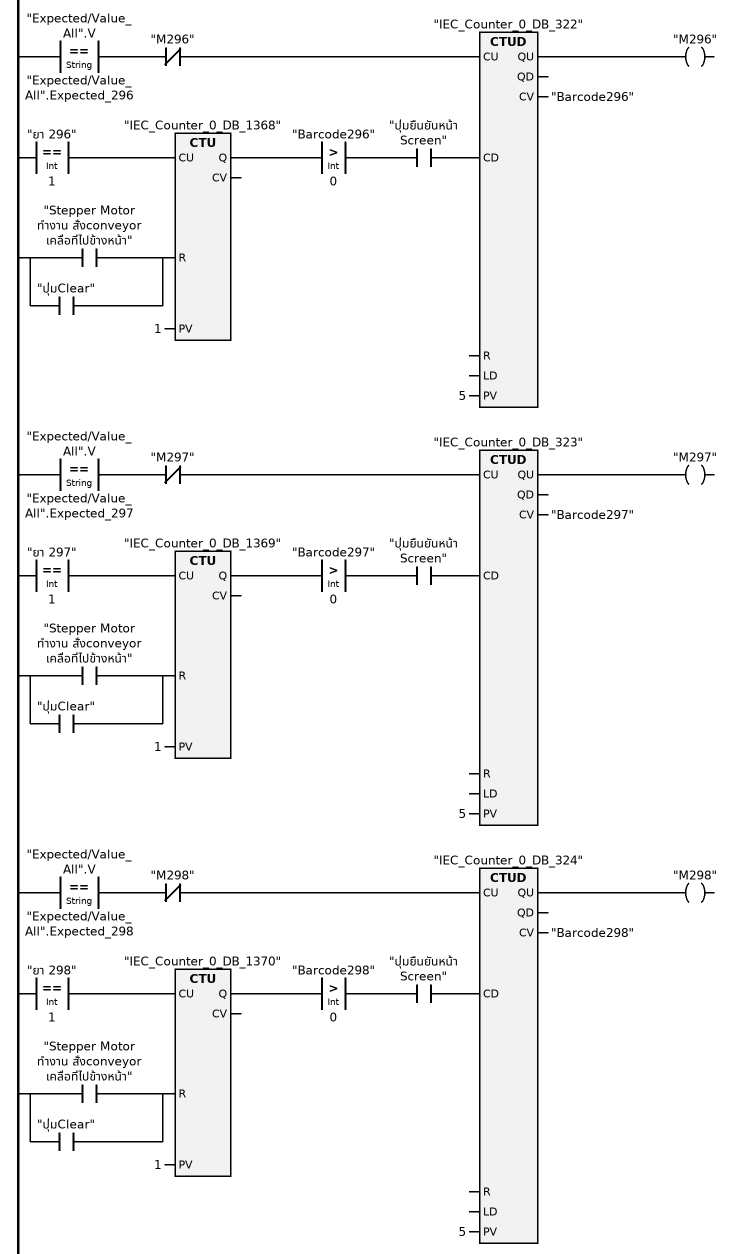
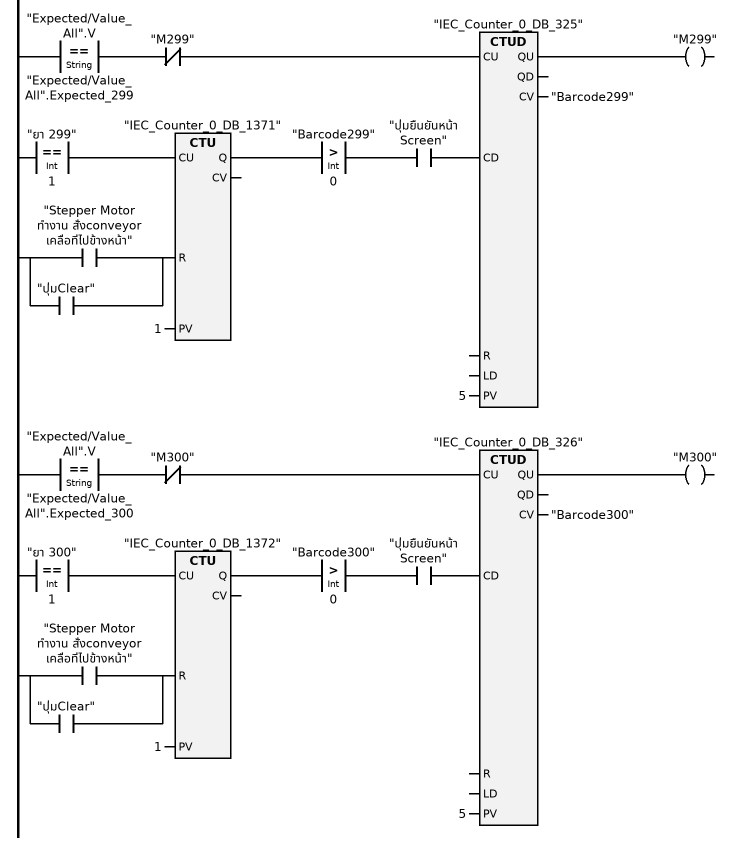
   "IEC_Counter_0_DB_1353".CTU(CU := "ยา 281" = 1,
                           R := "Stepper Motor ทำงาน สั่งconveyor เคลื่อที่ไปข้างหน้า" OR "ปุ่มClear",
                           PV := 1);
   "IEC_Counter_0_DB_307".CTUD(CU := ("Expected/Value_All".V = "Expected/Value_All".Expected_281) AND NOT "M281",
                           CD := "IEC_Counter_0_DB_1353".Q AND ("Barcode281" > 0) AND "ปุ่มยืนยันหน้า Screen",
                           PV := 5,
                           CV => "Barcode281");
   "M281" := "IEC_Counter_0_DB_307".QU;
   "IEC_Counter_0_DB_1354".CTU(CU := "ยา 282" = 1,
                           R := "Stepper Motor ทำงาน สั่งconveyor เคลื่อที่ไปข้างหน้า" OR "ปุ่มClear",
                           PV := 1);
   "IEC_Counter_0_DB_308".CTUD(CU := ("Expected/Value_All".V = "Expected/Value_All".Expected_282) AND NOT "M282",
                           CD := "IEC_Counter_0_DB_1354".Q AND ("Barcode282" > 0) AND "ปุ่มยืนยันหน้า Screen",
                           PV := 5,
                           CV => "Barcode282");
   "M282" := "IEC_Counter_0_DB_308".QU;
   "IEC_Counter_0_DB_1355".CTU(CU := "ยา 283" = 1,
                           R := "Stepper Motor ทำงาน สั่งconveyor เคลื่อที่ไปข้างหน้า" OR "ปุ่มClear",
                           PV := 1);
   "IEC_Counter_0_DB_309".CTUD(CU := ("Expected/Value_All".V = "Expected/Value_All".Expected_283) AND NOT "M283",
                           CD := "IEC_Counter_0_DB_1355".Q AND ("Barcode283" > 0) AND "ปุ่มยืนยันหน้า Screen",
                           PV := 5,
                           CV => "Barcode283");
   "M283" := "IEC_Counter_0_DB_309".QU;
   "IEC_Counter_0_DB_1356".CTU(CU := "ยา 284" = 1,
                           R := "Stepper Motor ทำงาน สั่งconveyor เคลื่อที่ไปข้างหน้า" OR "ปุ่มClear",
                           PV := 1);
   "IEC_Counter_0_DB_310".CTUD(CU := ("Expected/Value_All".V = "Expected/Value_All".Expected_284) AND NOT "M284",
                           CD := "IEC_Counter_0_DB_1356".Q AND ("Barcode284" > 0) AND "ปุ่มยืนยันหน้า Screen",
                           PV := 5,
                           CV => "Barcode284");
   "M284" := "IEC_Counter_0_DB_310".QU;
   "IEC_Counter_0_DB_1357".CTU(CU := "ยา 285" = 1,
                           R := "Stepper Motor ทำงาน สั่งconveyor เคลื่อที่ไปข้างหน้า" OR "ปุ่มClear",
                           PV := 1);
   "IEC_Counter_0_DB_311".CTUD(CU := ("Expected/Value_All".V = "Expected/Value_All".Expected_285) AND NOT "M285",
                           CD := "IEC_Counter_0_DB_1357".Q AND ("Barcode285" > 0) AND "ปุ่มยืนยันหน้า Screen",
                           PV := 5,
                           CV => "Barcode285");
   "M285" := "IEC_Counter_0_DB_311".QU;
   "IEC_Counter_0_DB_1358".CTU(CU := "ยา 286" = 1,
                           R := "Stepper Motor ทำงาน สั่งconveyor เคลื่อที่ไปข้างหน้า" OR "ปุ่มClear",
                           PV := 1);
   "IEC_Counter_0_DB_312".CTUD(CU := ("Expected/Value_All".V = "Expected/Value_All".Expected_286) AND NOT "M286",
                           CD := "IEC_Counter_0_DB_1358".Q AND ("Barcode286" > 0) AND "ปุ่มยืนยันหน้า Screen",
                           PV := 5,
                           CV => "Barcode286");
   "M286" := "IEC_Counter_0_DB_312".QU;
   "IEC_Counter_0_DB_1359".CTU(CU := "ยา 287" = 1,
                           R := "Stepper Motor ทำงาน สั่งconveyor เคลื่อที่ไปข้างหน้า" OR "ปุ่มClear",
                           PV := 1);
   "IEC_Counter_0_DB_313".CTUD(CU := ("Expected/Value_All".V = "Expected/Value_All".Expected_287) AND NOT "M287",
                           CD := "IEC_Counter_0_DB_1359".Q AND ("Barcode287" > 0) AND "ปุ่มยืนยันหน้า Screen",
                           PV := 5,
                           CV => "Barcode287");
   "M287" := "IEC_Counter_0_DB_313".QU;
   "IEC_Counter_0_DB_1360".CTU(CU := "ยา 288" = 1,
                           R := "Stepper Motor ทำงาน สั่งconveyor เคลื่อที่ไปข้างหน้า" OR "ปุ่มClear",
                           PV := 1);
   "IEC_Counter_0_DB_314".CTUD(CU := ("Expected/Value_All".V = "Expected/Value_All".Expected_288) AND NOT "M288",
                           CD := "IEC_Counter_0_DB_1360".Q AND ("Barcode288" > 0) AND "ปุ่มยืนยันหน้า Screen",
                           PV := 5,
                           CV => "Barcode288");
   "M288" := "IEC_Counter_0_DB_314".QU;
   "IEC_Counter_0_DB_1361".CTU(CU := "ยา 289" = 1,
                           R := "Stepper Motor ทำงาน สั่งconveyor เคลื่อที่ไปข้างหน้า" OR "ปุ่มClear",
                           PV := 1);
   "IEC_Counter_0_DB_315".CTUD(CU := ("Expected/Value_All".V = "Expected/Value_All".Expected_289) AND NOT "M289",
                           CD := "IEC_Counter_0_DB_1361".Q AND ("Barcode289" > 0) AND "ปุ่มยืนยันหน้า Screen",
                           PV := 5,
                           CV => "Barcode289");
   "M289" := "IEC_Counter_0_DB_315".QU;
   "IEC_Counter_0_DB_1362".CTU(CU := "ยา 290" = 1,
                           R := "Stepper Motor ทำงาน สั่งconveyor เคลื่อที่ไปข้างหน้า" OR "ปุ่มClear",
                           PV := 1);
   "IEC_Counter_0_DB_316".CTUD(CU := ("Expected/Value_All".V = "Expected/Value_All".Expected_290) AND NOT "M290",
                           CD := "IEC_Counter_0_DB_1362".Q AND ("Barcode290" > 0) AND "ปุ่มยืนยันหน้า Screen",
                           PV := 5,
                           CV => "Barcode290");
   "M290" := "IEC_Counter_0_DB_316".QU;
   "IEC_Counter_0_DB_1363".CTU(CU := "ยา 291" = 1,
                           R := "Stepper Motor ทำงาน สั่งconveyor เคลื่อที่ไปข้างหน้า" OR "ปุ่มClear",
                           PV := 1);
   "IEC_Counter_0_DB_317".CTUD(CU := ("Expected/Value_All".V = "Expected/Value_All".Expected_291) AND NOT "M291",
                           CD := "IEC_Counter_0_DB_1363".Q AND ("Barcode291" > 0) AND "ปุ่มยืนยันหน้า Screen",
                           PV := 5,
                           CV => "Barcode291");
   "M291" := "IEC_Counter_0_DB_317".QU;
   "IEC_Counter_0_DB_1364".CTU(CU := "ยา 292" = 1,
                           R := "Stepper Motor ทำงาน สั่งconveyor เคลื่อที่ไปข้างหน้า" OR "ปุ่มClear",
                           PV := 1);
   "IEC_Counter_0_DB_318".CTUD(CU := ("Expected/Value_All".V = "Expected/Value_All".Expected_292) AND NOT "M292",
                           CD := "IEC_Counter_0_DB_1364".Q AND ("Barcode292" > 0) AND "ปุ่มยืนยันหน้า Screen",
                           PV := 5,
                           CV => "Barcode292");
   "M292" := "IEC_Counter_0_DB_318".QU;
   "IEC_Counter_0_DB_1365".CTU(CU := "ยา 293" = 1,
                           R := "Stepper Motor ทำงาน สั่งconveyor เคลื่อที่ไปข้างหน้า" OR "ปุ่มClear",
                           PV := 1);
   "IEC_Counter_0_DB_319".CTUD(CU := ("Expected/Value_All".V = "Expected/Value_All".Expected_293) AND NOT "M293",
                           CD := "IEC_Counter_0_DB_1365".Q AND ("Barcode293" > 0) AND "ปุ่มยืนยันหน้า Screen",
                           PV := 5,
                           CV => "Barcode293");
   "M293" := "IEC_Counter_0_DB_319".QU;
   "IEC_Counter_0_DB_1366".CTU(CU := "ยา 294" = 1,
                           R := "Stepper Motor ทำงาน สั่งconveyor เคลื่อที่ไปข้างหน้า" OR "ปุ่มClear",
                           PV := 1);
   "IEC_Counter_0_DB_320".CTUD(CU := ("Expected/Value_All".V = "Expected/Value_All".Expected_294) AND NOT "M294",
                           CD := "IEC_Counter_0_DB_1366".Q AND ("Barcode294" > 0) AND "ปุ่มยืนยันหน้า Screen",
                           PV := 5,
                           CV => "Barcode294");
   "M294" := "IEC_Counter_0_DB_320".QU;
   "IEC_Counter_0_DB_1367".CTU(CU := "ยา 295" = 1,
                           R := "Stepper Motor ทำงาน สั่งconveyor เคลื่อที่ไปข้างหน้า" OR "ปุ่มClear",
                           PV := 1);
   "IEC_Counter_0_DB_321".CTUD(CU := ("Expected/Value_All".V = "Expected/Value_All".Expected_295) AND NOT "M295",
                           CD := "IEC_Counter_0_DB_1367".Q AND ("Barcode295" > 0) AND "ปุ่มยืนยันหน้า Screen",
                           PV := 5,
                           CV => "Barcode295");
   "M295" := "IEC_Counter_0_DB_321".QU;
   "IEC_Counter_0_DB_1368".CTU(CU := "ยา 296" = 1,
                           R := "Stepper Motor ทำงาน สั่งconveyor เคลื่อที่ไปข้างหน้า" OR "ปุ่มClear",
                           PV := 1);
   "IEC_Counter_0_DB_322".CTUD(CU := ("Expected/Value_All".V = "Expected/Value_All".Expected_296) AND NOT "M296",
                           CD := "IEC_Counter_0_DB_1368".Q AND ("Barcode296" > 0) AND "ปุ่มยืนยันหน้า Screen",
                           PV := 5,
                           CV => "Barcode296");
   "M296" := "IEC_Counter_0_DB_322".QU;
   "IEC_Counter_0_DB_1369".CTU(CU := "ยา 297" = 1,
                           R := "Stepper Motor ทำงาน สั่งconveyor เคลื่อที่ไปข้างหน้า" OR "ปุ่มClear",
                           PV := 1);
   "IEC_Counter_0_DB_323".CTUD(CU := ("Expected/Value_All".V = "Expected/Value_All".Expected_297) AND NOT "M297",
                           CD := "IEC_Counter_0_DB_1369".Q AND ("Barcode297" > 0) AND "ปุ่มยืนยันหน้า Screen",
                           PV := 5,
                           CV => "Barcode297");
   "M297" := "IEC_Counter_0_DB_323".QU;
   "IEC_Counter_0_DB_1370".CTU(CU := "ยา 298" = 1,
                           R := "Stepper Motor ทำงาน สั่งconveyor เคลื่อที่ไปข้างหน้า" OR "ปุ่มClear",
                           PV := 1);
   "IEC_Counter_0_DB_324".CTUD(CU := ("Expected/Value_All".V = "Expected/Value_All".Expected_298) AND NOT "M298",
                           CD := "IEC_Counter_0_DB_1370".Q AND ("Barcode298" > 0) AND "ปุ่มยืนยันหน้า Screen",
                           PV := 5,
                           CV => "Barcode298");
   "M298" := "IEC_Counter_0_DB_324".QU;
   "IEC_Counter_0_DB_1371".CTU(CU := "ยา 299" = 1,
                           R := "Stepper Motor ทำงาน สั่งconveyor เคลื่อที่ไปข้างหน้า" OR "ปุ่มClear",
                           PV := 1);
   "IEC_Counter_0_DB_325".CTUD(CU := ("Expected/Value_All".V = "Expected/Value_All".Expected_299) AND NOT "M299",
                           CD := "IEC_Counter_0_DB_1371".Q AND ("Barcode299" > 0) AND "ปุ่มยืนยันหน้า Screen",
                           PV := 5,
                           CV => "Barcode299");
   "M299" := "IEC_Counter_0_DB_325".QU;
   "IEC_Counter_0_DB_1372".CTU(CU := "ยา 300" = 1,
                           R := "Stepper Motor ทำงาน สั่งconveyor เคลื่อที่ไปข้างหน้า" OR "ปุ่มClear",
                           PV := 1);
   "IEC_Counter_0_DB_326".CTUD(CU := ("Expected/Value_All".V = "Expected/Value_All".Expected_300) AND NOT "M300",
                           CD := "IEC_Counter_0_DB_1372".Q AND ("Barcode300" > 0) AND "ปุ่มยืนยันหน้า Screen",
                           PV := 5,
                           CV => "Barcode300");
   "M300" := "IEC_Counter_0_DB_326".QU;
END_REGION

REGION Network 16
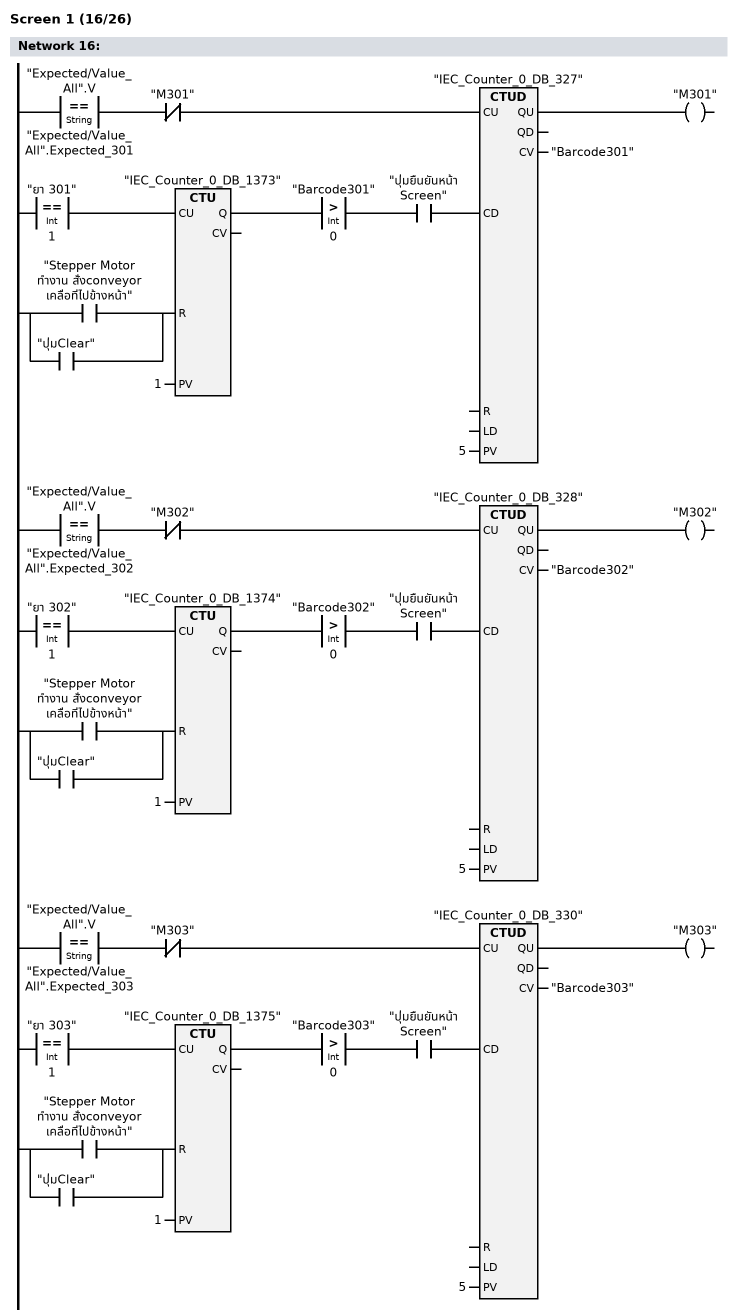
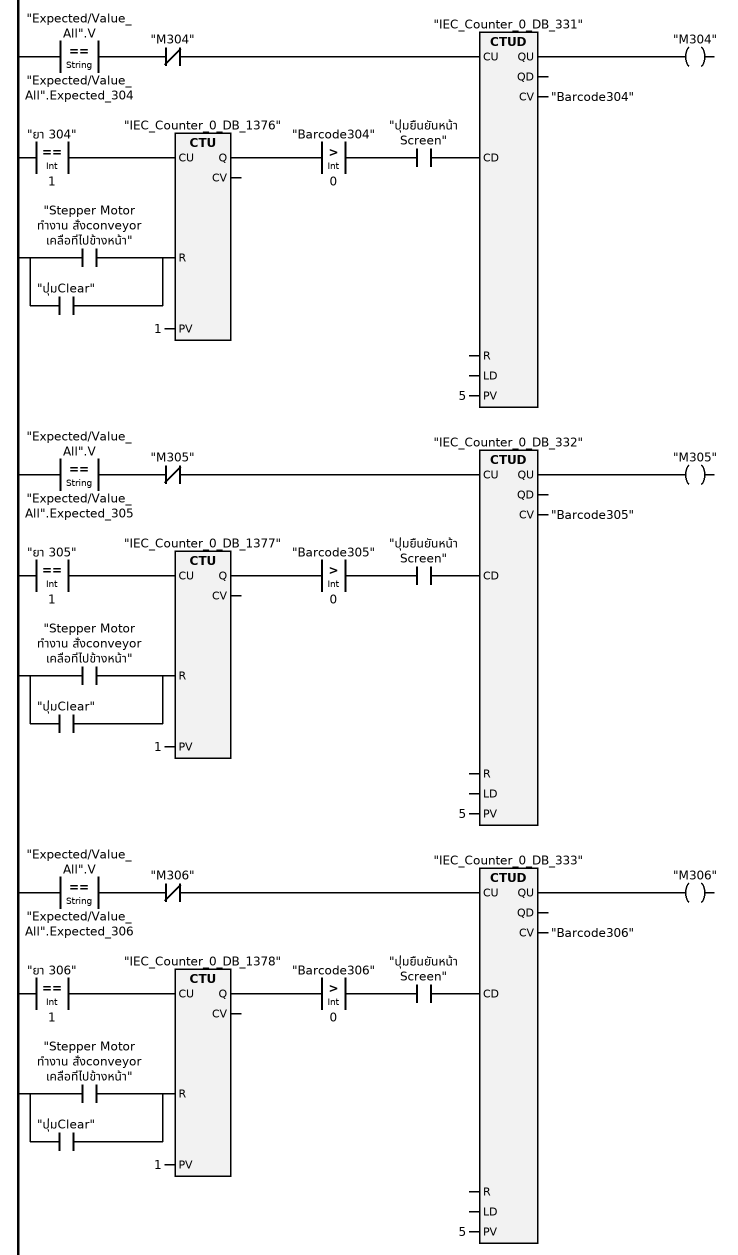
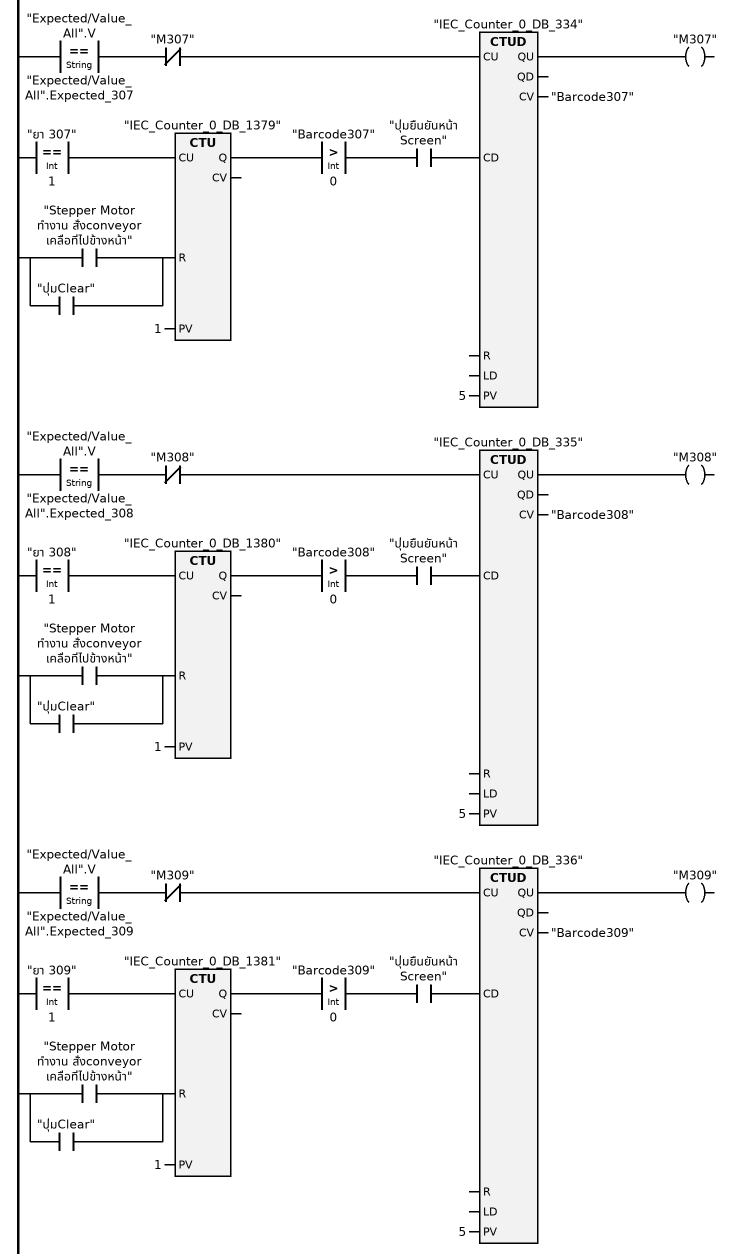
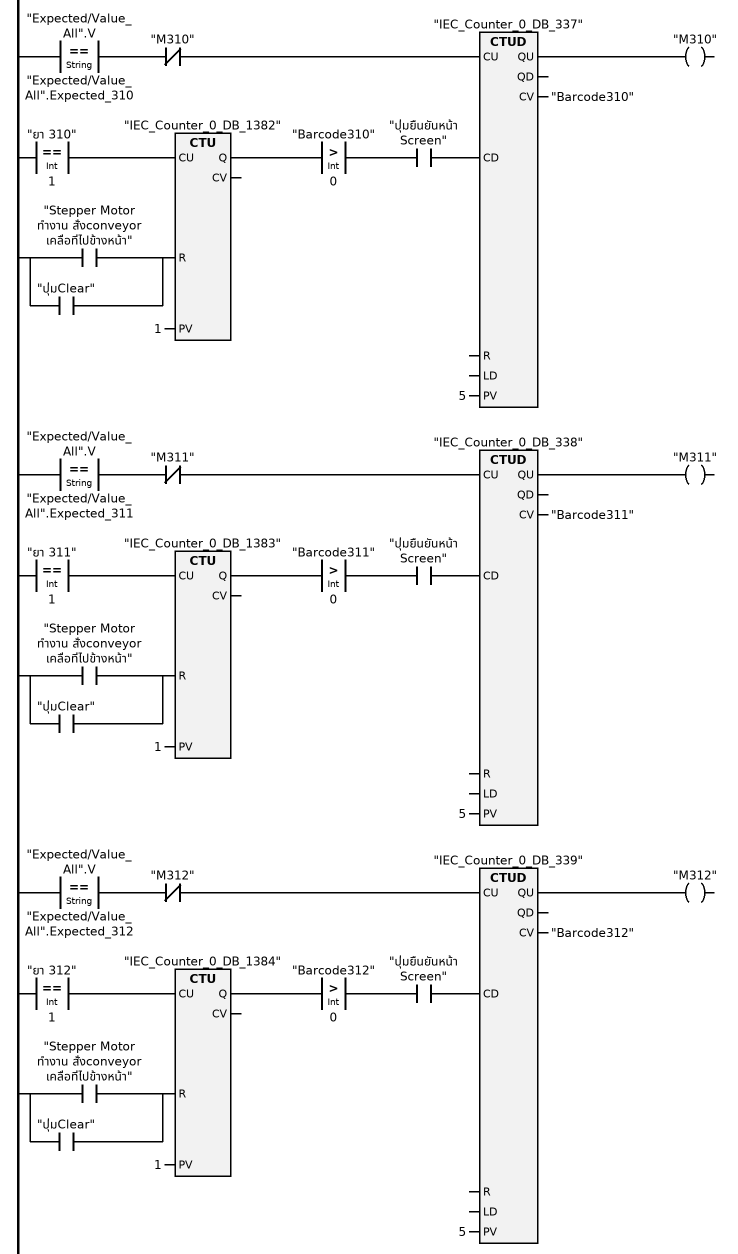
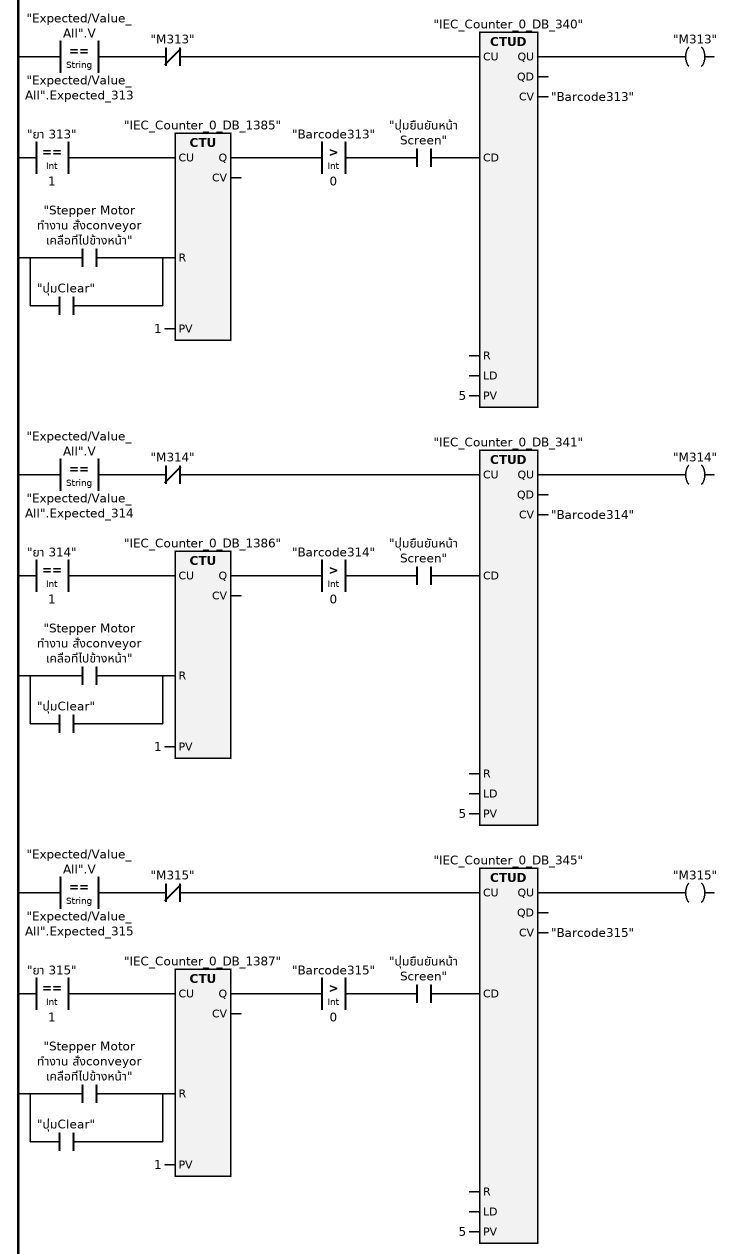
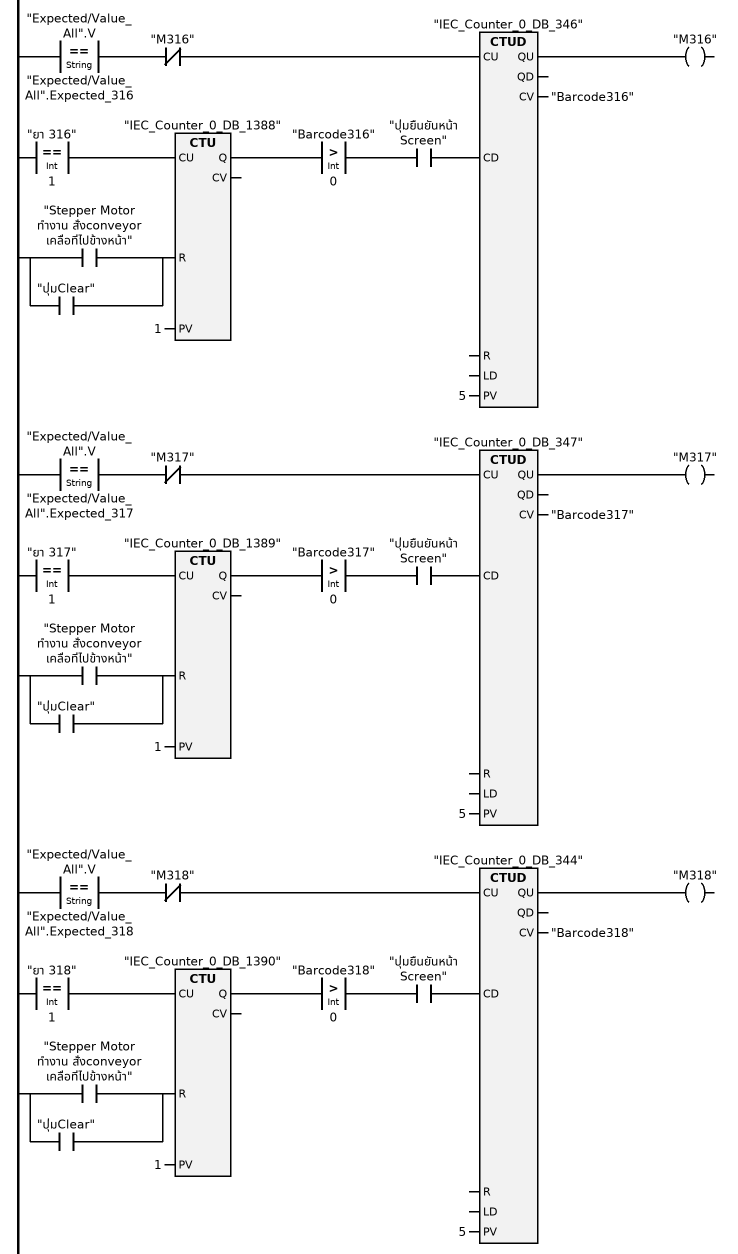
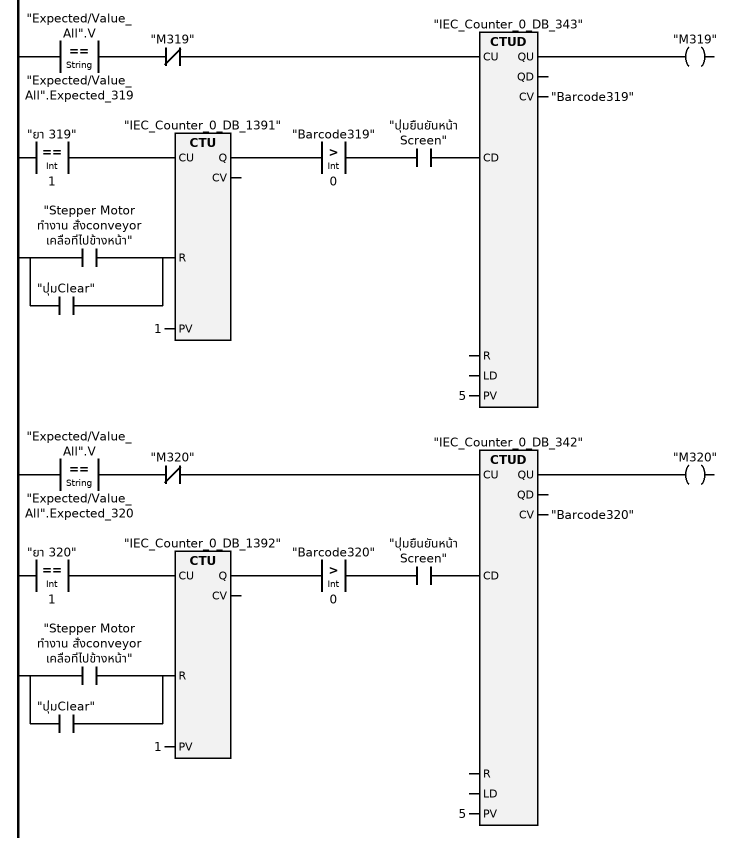
   "IEC_Counter_0_DB_1373".CTU(CU := "ยา 301" = 1,
                           R := "Stepper Motor ทำงาน สั่งconveyor เคลื่อที่ไปข้างหน้า" OR "ปุ่มClear",
                           PV := 1);
   "IEC_Counter_0_DB_327".CTUD(CU := ("Expected/Value_All".V = "Expected/Value_All".Expected_301) AND NOT "M301",
                           CD := "IEC_Counter_0_DB_1373".Q AND ("Barcode301" > 0) AND "ปุ่มยืนยันหน้า Screen",
                           PV := 5,
                           CV => "Barcode301");
   "M301" := "IEC_Counter_0_DB_327".QU;
   "IEC_Counter_0_DB_1374".CTU(CU := "ยา 302" = 1,
                           R := "Stepper Motor ทำงาน สั่งconveyor เคลื่อที่ไปข้างหน้า" OR "ปุ่มClear",
                           PV := 1);
   "IEC_Counter_0_DB_328".CTUD(CU := ("Expected/Value_All".V = "Expected/Value_All".Expected_302) AND NOT "M302",
                           CD := "IEC_Counter_0_DB_1374".Q AND ("Barcode302" > 0) AND "ปุ่มยืนยันหน้า Screen",
                           PV := 5,
                           CV => "Barcode302");
   "M302" := "IEC_Counter_0_DB_328".QU;
   "IEC_Counter_0_DB_1375".CTU(CU := "ยา 303" = 1,
                           R := "Stepper Motor ทำงาน สั่งconveyor เคลื่อที่ไปข้างหน้า" OR "ปุ่มClear",
                           PV := 1);
   "IEC_Counter_0_DB_330".CTUD(CU := ("Expected/Value_All".V = "Expected/Value_All".Expected_303) AND NOT "M303",
                           CD := "IEC_Counter_0_DB_1375".Q AND ("Barcode303" > 0) AND "ปุ่มยืนยันหน้า Screen",
                           PV := 5,
                           CV => "Barcode303");
   "M303" := "IEC_Counter_0_DB_330".QU;
   "IEC_Counter_0_DB_1376".CTU(CU := "ยา 304" = 1,
                           R := "Stepper Motor ทำงาน สั่งconveyor เคลื่อที่ไปข้างหน้า" OR "ปุ่มClear",
                           PV := 1);
   "IEC_Counter_0_DB_331".CTUD(CU := ("Expected/Value_All".V = "Expected/Value_All".Expected_304) AND NOT "M304",
                           CD := "IEC_Counter_0_DB_1376".Q AND ("Barcode304" > 0) AND "ปุ่มยืนยันหน้า Screen",
                           PV := 5,
                           CV => "Barcode304");
   "M304" := "IEC_Counter_0_DB_331".QU;
   "IEC_Counter_0_DB_1377".CTU(CU := "ยา 305" = 1,
                           R := "Stepper Motor ทำงาน สั่งconveyor เคลื่อที่ไปข้างหน้า" OR "ปุ่มClear",
                           PV := 1);
   "IEC_Counter_0_DB_332".CTUD(CU := ("Expected/Value_All".V = "Expected/Value_All".Expected_305) AND NOT "M305",
                           CD := "IEC_Counter_0_DB_1377".Q AND ("Barcode305" > 0) AND "ปุ่มยืนยันหน้า Screen",
                           PV := 5,
                           CV => "Barcode305");
   "M305" := "IEC_Counter_0_DB_332".QU;
   "IEC_Counter_0_DB_1378".CTU(CU := "ยา 306" = 1,
                           R := "Stepper Motor ทำงาน สั่งconveyor เคลื่อที่ไปข้างหน้า" OR "ปุ่มClear",
                           PV := 1);
   "IEC_Counter_0_DB_333".CTUD(CU := ("Expected/Value_All".V = "Expected/Value_All".Expected_306) AND NOT "M306",
                           CD := "IEC_Counter_0_DB_1378".Q AND ("Barcode306" > 0) AND "ปุ่มยืนยันหน้า Screen",
                           PV := 5,
                           CV => "Barcode306");
   "M306" := "IEC_Counter_0_DB_333".QU;
   "IEC_Counter_0_DB_1379".CTU(CU := "ยา 307" = 1,
                           R := "Stepper Motor ทำงาน สั่งconveyor เคลื่อที่ไปข้างหน้า" OR "ปุ่มClear",
                           PV := 1);
   "IEC_Counter_0_DB_334".CTUD(CU := ("Expected/Value_All".V = "Expected/Value_All".Expected_307) AND NOT "M307",
                           CD := "IEC_Counter_0_DB_1379".Q AND ("Barcode307" > 0) AND "ปุ่มยืนยันหน้า Screen",
                           PV := 5,
                           CV => "Barcode307");
   "M307" := "IEC_Counter_0_DB_334".QU;
   "IEC_Counter_0_DB_1380".CTU(CU := "ยา 308" = 1,
                           R := "Stepper Motor ทำงาน สั่งconveyor เคลื่อที่ไปข้างหน้า" OR "ปุ่มClear",
                           PV := 1);
   "IEC_Counter_0_DB_335".CTUD(CU := ("Expected/Value_All".V = "Expected/Value_All".Expected_308) AND NOT "M308",
                           CD := "IEC_Counter_0_DB_1380".Q AND ("Barcode308" > 0) AND "ปุ่มยืนยันหน้า Screen",
                           PV := 5,
                           CV => "Barcode308");
   "M308" := "IEC_Counter_0_DB_335".QU;
   "IEC_Counter_0_DB_1381".CTU(CU := "ยา 309" = 1,
                           R := "Stepper Motor ทำงาน สั่งconveyor เคลื่อที่ไปข้างหน้า" OR "ปุ่มClear",
                           PV := 1);
   "IEC_Counter_0_DB_336".CTUD(CU := ("Expected/Value_All".V = "Expected/Value_All".Expected_309) AND NOT "M309",
                           CD := "IEC_Counter_0_DB_1381".Q AND ("Barcode309" > 0) AND "ปุ่มยืนยันหน้า Screen",
                           PV := 5,
                           CV => "Barcode309");
   "M309" := "IEC_Counter_0_DB_336".QU;
   "IEC_Counter_0_DB_1382".CTU(CU := "ยา 310" = 1,
                           R := "Stepper Motor ทำงาน สั่งconveyor เคลื่อที่ไปข้างหน้า" OR "ปุ่มClear",
                           PV := 1);
   "IEC_Counter_0_DB_337".CTUD(CU := ("Expected/Value_All".V = "Expected/Value_All".Expected_310) AND NOT "M310",
                           CD := "IEC_Counter_0_DB_1382".Q AND ("Barcode310" > 0) AND "ปุ่มยืนยันหน้า Screen",
                           PV := 5,
                           CV => "Barcode310");
   "M310" := "IEC_Counter_0_DB_337".QU;
   "IEC_Counter_0_DB_1383".CTU(CU := "ยา 311" = 1,
                           R := "Stepper Motor ทำงาน สั่งconveyor เคลื่อที่ไปข้างหน้า" OR "ปุ่มClear",
                           PV := 1);
   "IEC_Counter_0_DB_338".CTUD(CU := ("Expected/Value_All".V = "Expected/Value_All".Expected_311) AND NOT "M311",
                           CD := "IEC_Counter_0_DB_1383".Q AND ("Barcode311" > 0) AND "ปุ่มยืนยันหน้า Screen",
                           PV := 5,
                           CV => "Barcode311");
   "M311" := "IEC_Counter_0_DB_338".QU;
   "IEC_Counter_0_DB_1384".CTU(CU := "ยา 312" = 1,
                           R := "Stepper Motor ทำงาน สั่งconveyor เคลื่อที่ไปข้างหน้า" OR "ปุ่มClear",
                           PV := 1);
   "IEC_Counter_0_DB_339".CTUD(CU := ("Expected/Value_All".V = "Expected/Value_All".Expected_312) AND NOT "M312",
                           CD := "IEC_Counter_0_DB_1384".Q AND ("Barcode312" > 0) AND "ปุ่มยืนยันหน้า Screen",
                           PV := 5,
                           CV => "Barcode312");
   "M312" := "IEC_Counter_0_DB_339".QU;
   "IEC_Counter_0_DB_1385".CTU(CU := "ยา 313" = 1,
                           R := "Stepper Motor ทำงาน สั่งconveyor เคลื่อที่ไปข้างหน้า" OR "ปุ่มClear",
                           PV := 1);
   "IEC_Counter_0_DB_340".CTUD(CU := ("Expected/Value_All".V = "Expected/Value_All".Expected_313) AND NOT "M313",
                           CD := "IEC_Counter_0_DB_1385".Q AND ("Barcode313" > 0) AND "ปุ่มยืนยันหน้า Screen",
                           PV := 5,
                           CV => "Barcode313");
   "M313" := "IEC_Counter_0_DB_340".QU;
   "IEC_Counter_0_DB_1386".CTU(CU := "ยา 314" = 1,
                           R := "Stepper Motor ทำงาน สั่งconveyor เคลื่อที่ไปข้างหน้า" OR "ปุ่มClear",
                           PV := 1);
   "IEC_Counter_0_DB_341".CTUD(CU := ("Expected/Value_All".V = "Expected/Value_All".Expected_314) AND NOT "M314",
                           CD := "IEC_Counter_0_DB_1386".Q AND ("Barcode314" > 0) AND "ปุ่มยืนยันหน้า Screen",
                           PV := 5,
                           CV => "Barcode314");
   "M314" := "IEC_Counter_0_DB_341".QU;
   "IEC_Counter_0_DB_1387".CTU(CU := "ยา 315" = 1,
                           R := "Stepper Motor ทำงาน สั่งconveyor เคลื่อที่ไปข้างหน้า" OR "ปุ่มClear",
                           PV := 1);
   "IEC_Counter_0_DB_345".CTUD(CU := ("Expected/Value_All".V = "Expected/Value_All".Expected_315) AND NOT "M315",
                           CD := "IEC_Counter_0_DB_1387".Q AND ("Barcode315" > 0) AND "ปุ่มยืนยันหน้า Screen",
                           PV := 5,
                           CV => "Barcode315");
   "M315" := "IEC_Counter_0_DB_345".QU;
   "IEC_Counter_0_DB_1388".CTU(CU := "ยา 316" = 1,
                           R := "Stepper Motor ทำงาน สั่งconveyor เคลื่อที่ไปข้างหน้า" OR "ปุ่มClear",
                           PV := 1);
   "IEC_Counter_0_DB_346".CTUD(CU := ("Expected/Value_All".V = "Expected/Value_All".Expected_316) AND NOT "M316",
                           CD := "IEC_Counter_0_DB_1388".Q AND ("Barcode316" > 0) AND "ปุ่มยืนยันหน้า Screen",
                           PV := 5,
                           CV => "Barcode316");
   "M316" := "IEC_Counter_0_DB_346".QU;
   "IEC_Counter_0_DB_1389".CTU(CU := "ยา 317" = 1,
                           R := "Stepper Motor ทำงาน สั่งconveyor เคลื่อที่ไปข้างหน้า" OR "ปุ่มClear",
                           PV := 1);
   "IEC_Counter_0_DB_347".CTUD(CU := ("Expected/Value_All".V = "Expected/Value_All".Expected_317) AND NOT "M317",
                           CD := "IEC_Counter_0_DB_1389".Q AND ("Barcode317" > 0) AND "ปุ่มยืนยันหน้า Screen",
                           PV := 5,
                           CV => "Barcode317");
   "M317" := "IEC_Counter_0_DB_347".QU;
   "IEC_Counter_0_DB_1390".CTU(CU := "ยา 318" = 1,
                           R := "Stepper Motor ทำงาน สั่งconveyor เคลื่อที่ไปข้างหน้า" OR "ปุ่มClear",
                           PV := 1);
   "IEC_Counter_0_DB_344".CTUD(CU := ("Expected/Value_All".V = "Expected/Value_All".Expected_318) AND NOT "M318",
                           CD := "IEC_Counter_0_DB_1390".Q AND ("Barcode318" > 0) AND "ปุ่มยืนยันหน้า Screen",
                           PV := 5,
                           CV => "Barcode318");
   "M318" := "IEC_Counter_0_DB_344".QU;
   "IEC_Counter_0_DB_1391".CTU(CU := "ยา 319" = 1,
                           R := "Stepper Motor ทำงาน สั่งconveyor เคลื่อที่ไปข้างหน้า" OR "ปุ่มClear",
                           PV := 1);
   "IEC_Counter_0_DB_343".CTUD(CU := ("Expected/Value_All".V = "Expected/Value_All".Expected_319) AND NOT "M319",
                           CD := "IEC_Counter_0_DB_1391".Q AND ("Barcode319" > 0) AND "ปุ่มยืนยันหน้า Screen",
                           PV := 5,
                           CV => "Barcode319");
   "M319" := "IEC_Counter_0_DB_343".QU;
   "IEC_Counter_0_DB_1392".CTU(CU := "ยา 320" = 1,
                           R := "Stepper Motor ทำงาน สั่งconveyor เคลื่อที่ไปข้างหน้า" OR "ปุ่มClear",
                           PV := 1);
   "IEC_Counter_0_DB_342".CTUD(CU := ("Expected/Value_All".V = "Expected/Value_All".Expected_320) AND NOT "M320",
                           CD := "IEC_Counter_0_DB_1392".Q AND ("Barcode320" > 0) AND "ปุ่มยืนยันหน้า Screen",
                           PV := 5,
                           CV => "Barcode320");
   "M320" := "IEC_Counter_0_DB_342".QU;
END_REGION

REGION Network 17
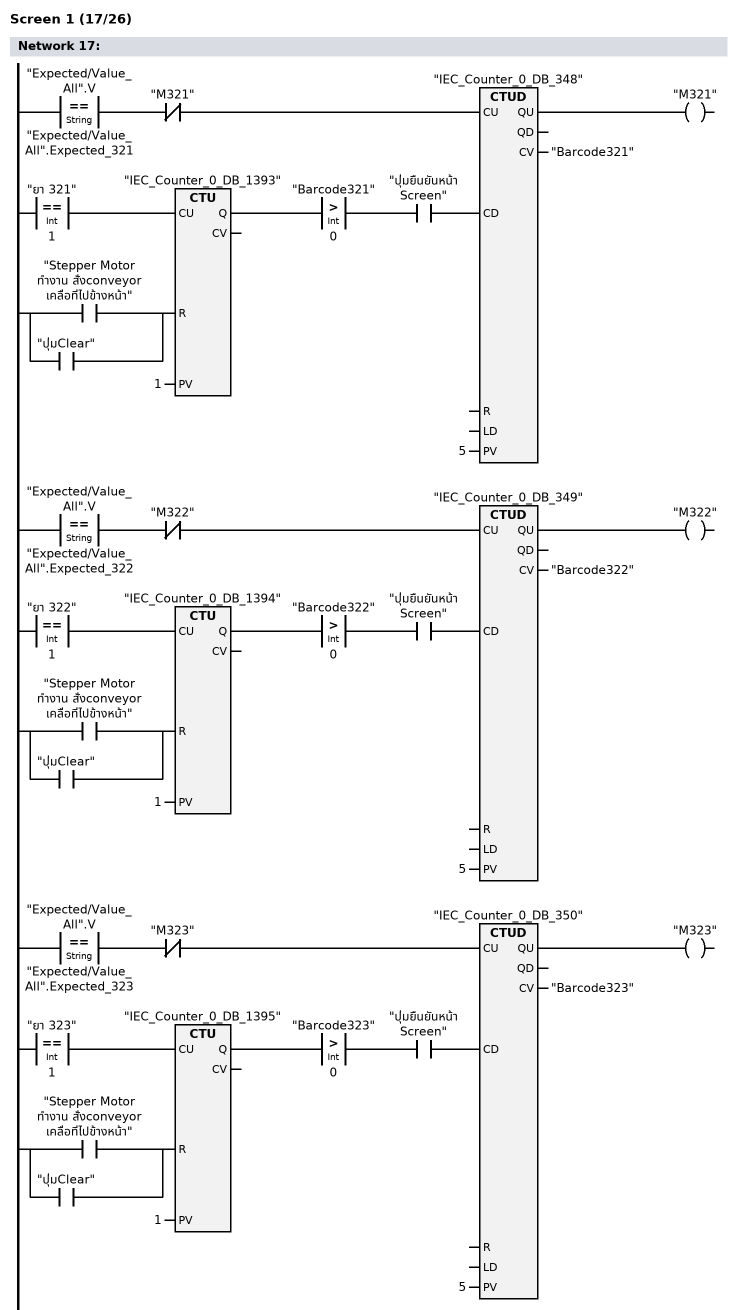
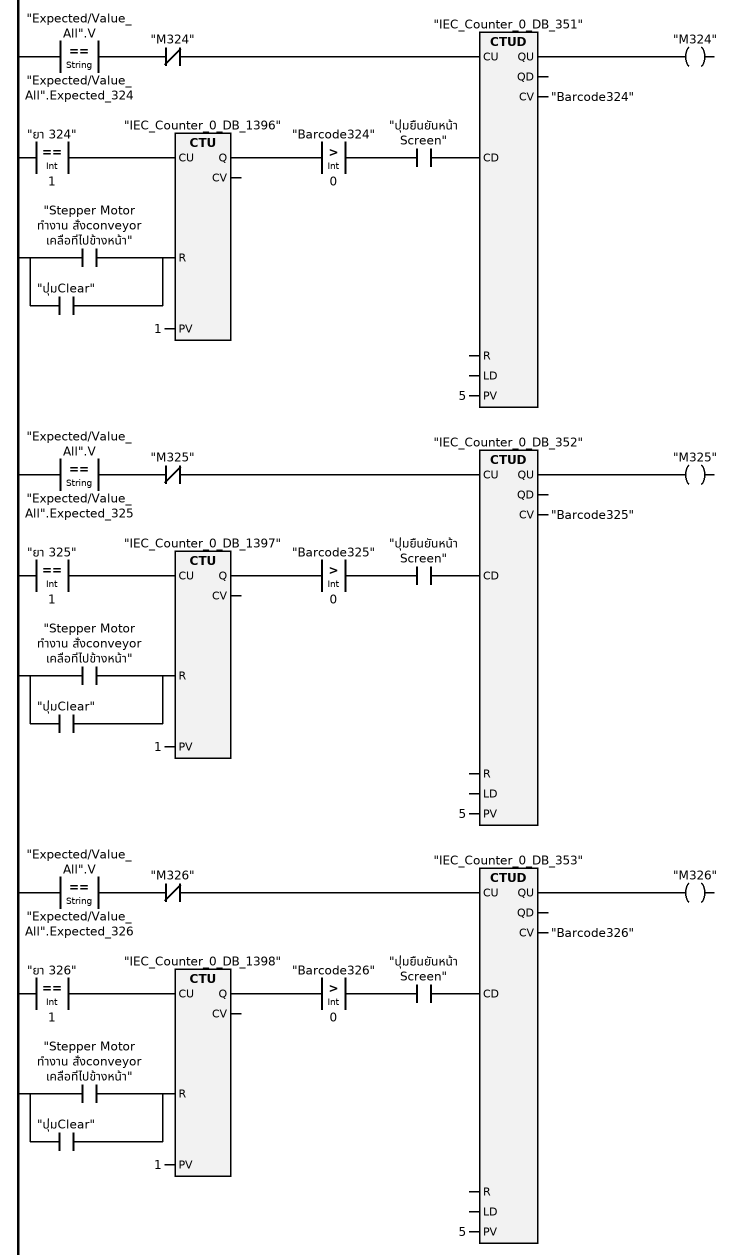
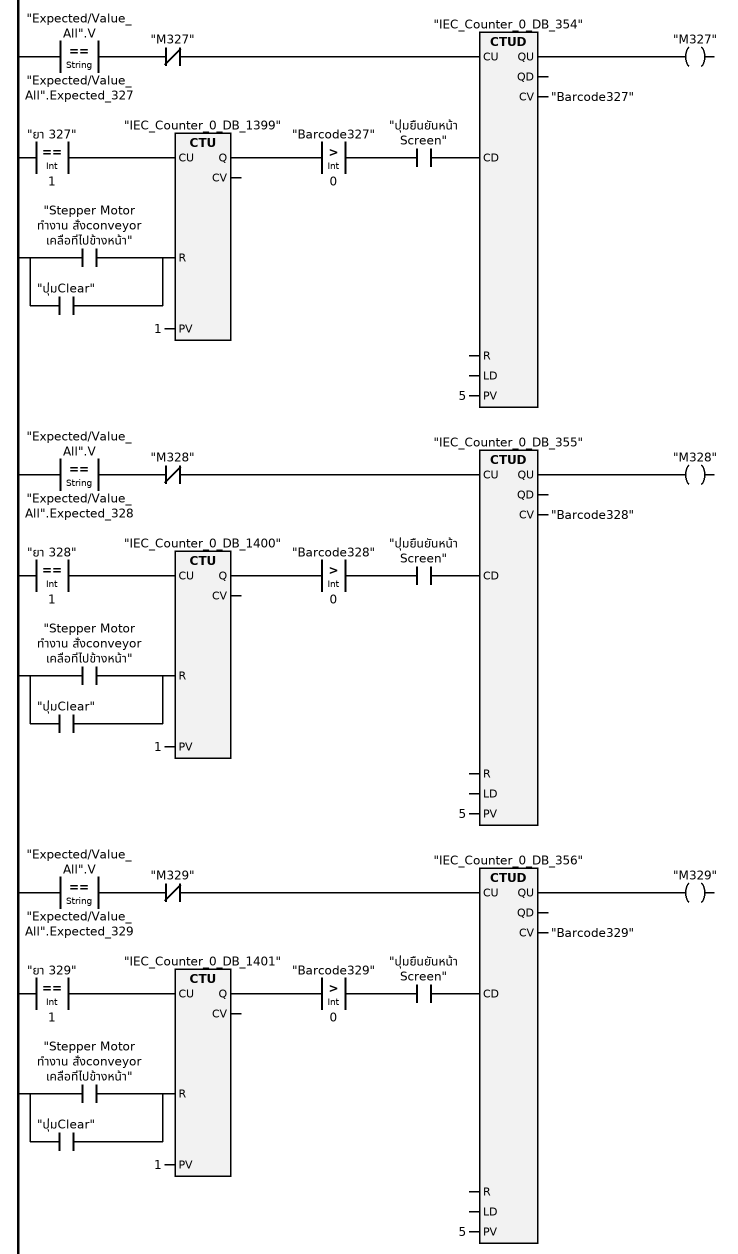
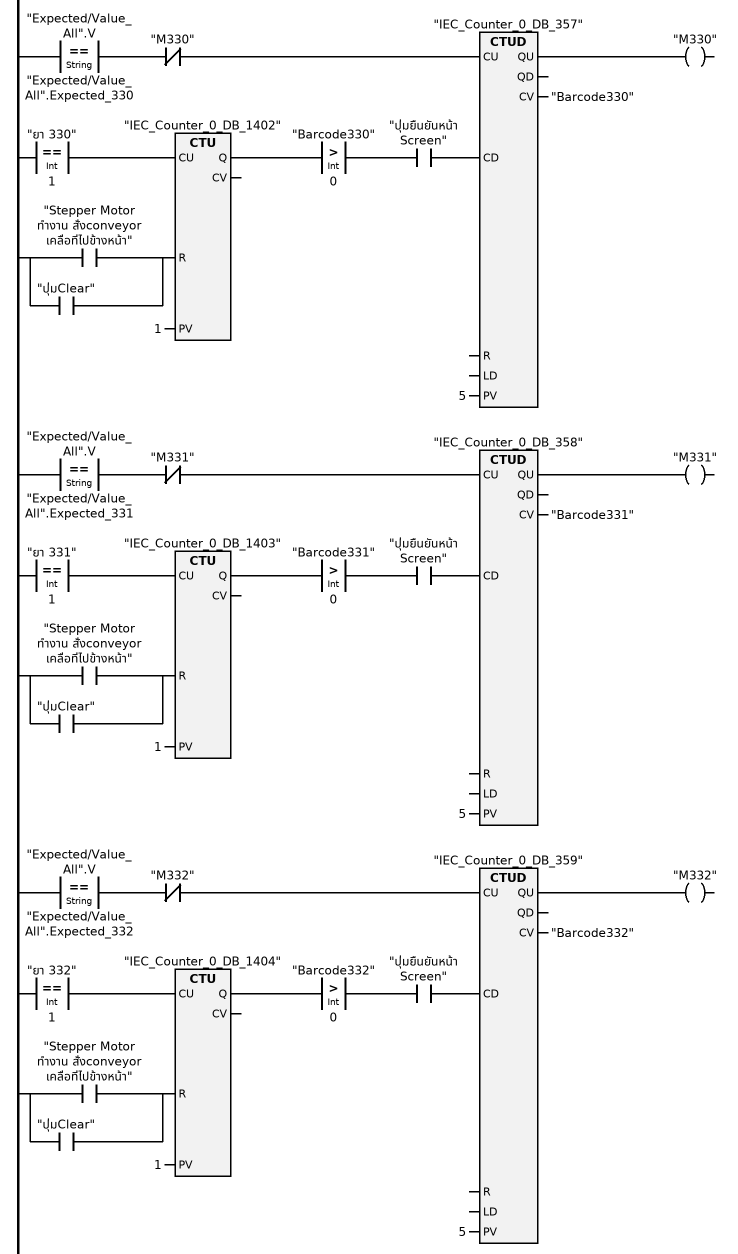
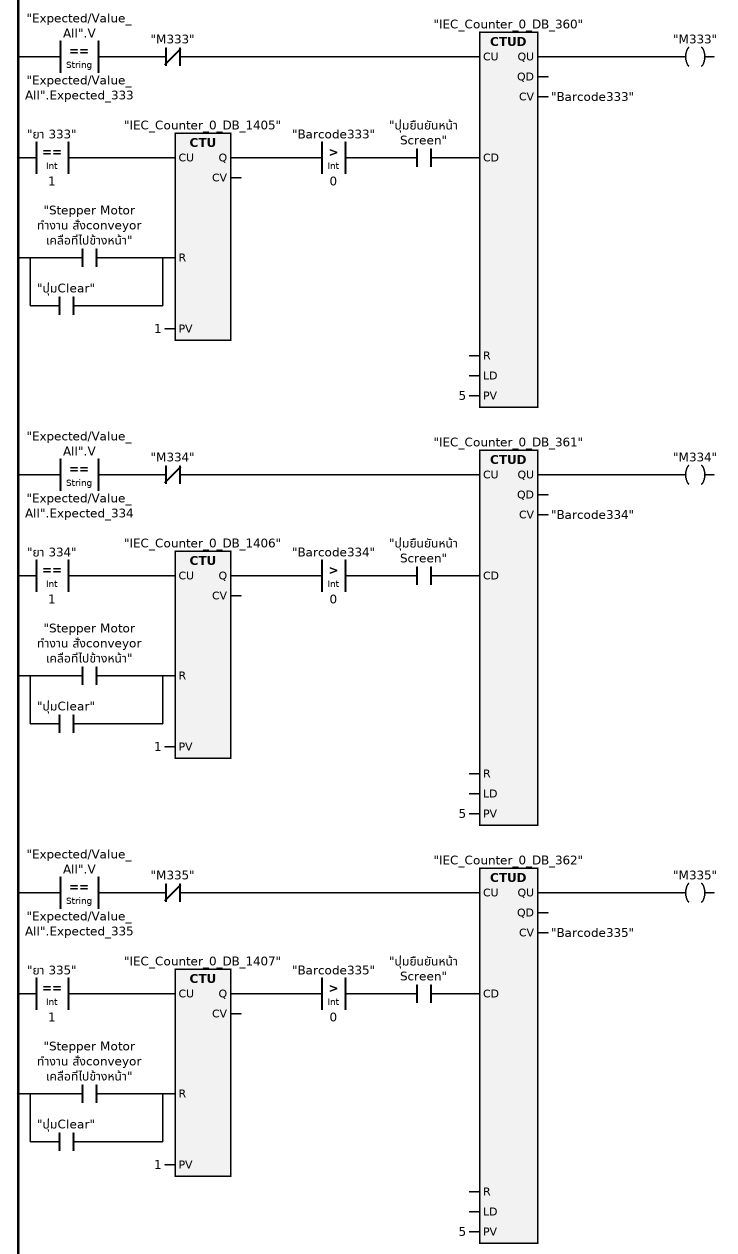
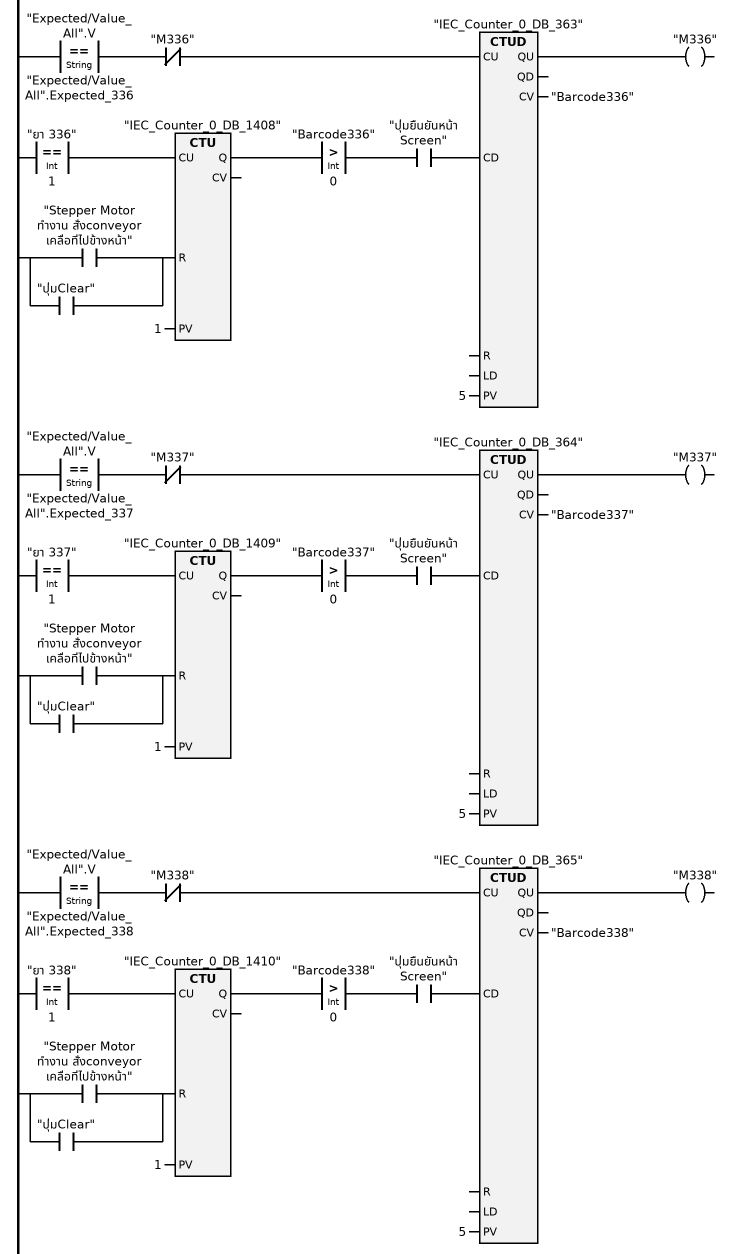
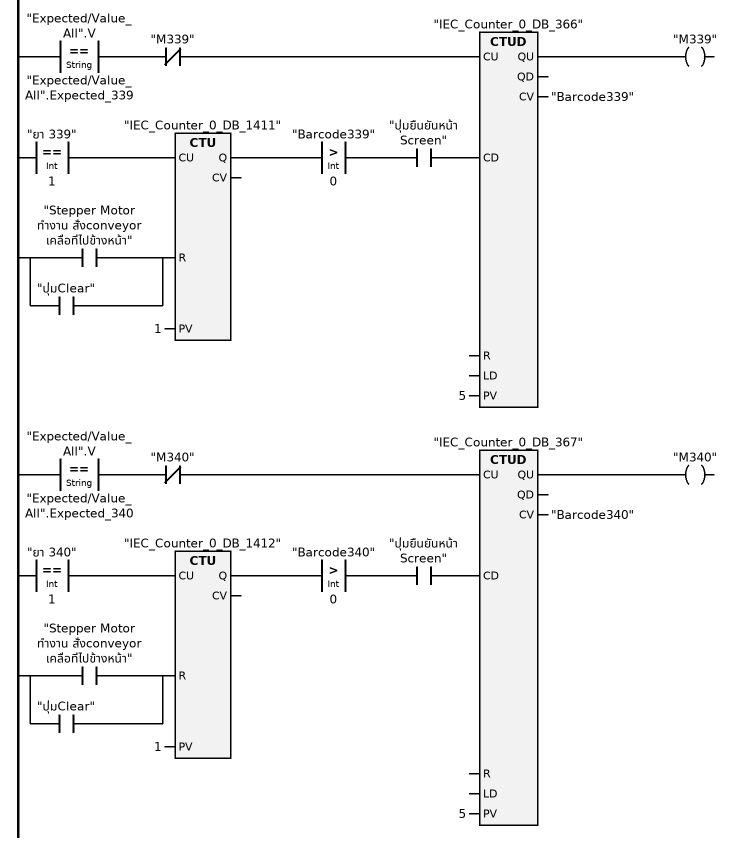
   "IEC_Counter_0_DB_1393".CTU(CU := "ยา 321" = 1,
                           R := "Stepper Motor ทำงาน สั่งconveyor เคลื่อที่ไปข้างหน้า" OR "ปุ่มClear",
                           PV := 1);
   "IEC_Counter_0_DB_348".CTUD(CU := ("Expected/Value_All".V = "Expected/Value_All".Expected_321) AND NOT "M321",
                           CD := "IEC_Counter_0_DB_1393".Q AND ("Barcode321" > 0) AND "ปุ่มยืนยันหน้า Screen",
                           PV := 5,
                           CV => "Barcode321");
   "M321" := "IEC_Counter_0_DB_348".QU;
   "IEC_Counter_0_DB_1394".CTU(CU := "ยา 322" = 1,
                           R := "Stepper Motor ทำงาน สั่งconveyor เคลื่อที่ไปข้างหน้า" OR "ปุ่มClear",
                           PV := 1);
   "IEC_Counter_0_DB_349".CTUD(CU := ("Expected/Value_All".V = "Expected/Value_All".Expected_322) AND NOT "M322",
                           CD := "IEC_Counter_0_DB_1394".Q AND ("Barcode322" > 0) AND "ปุ่มยืนยันหน้า Screen",
                           PV := 5,
                           CV => "Barcode322");
   "M322" := "IEC_Counter_0_DB_349".QU;
   "IEC_Counter_0_DB_1395".CTU(CU := "ยา 323" = 1,
                           R := "Stepper Motor ทำงาน สั่งconveyor เคลื่อที่ไปข้างหน้า" OR "ปุ่มClear",
                           PV := 1);
   "IEC_Counter_0_DB_350".CTUD(CU := ("Expected/Value_All".V = "Expected/Value_All".Expected_323) AND NOT "M323",
                           CD := "IEC_Counter_0_DB_1395".Q AND ("Barcode323" > 0) AND "ปุ่มยืนยันหน้า Screen",
                           PV := 5,
                           CV => "Barcode323");
   "M323" := "IEC_Counter_0_DB_350".QU;
   "IEC_Counter_0_DB_1396".CTU(CU := "ยา 324" = 1,
                           R := "Stepper Motor ทำงาน สั่งconveyor เคลื่อที่ไปข้างหน้า" OR "ปุ่มClear",
                           PV := 1);
   "IEC_Counter_0_DB_351".CTUD(CU := ("Expected/Value_All".V = "Expected/Value_All".Expected_324) AND NOT "M324",
                           CD := "IEC_Counter_0_DB_1396".Q AND ("Barcode324" > 0) AND "ปุ่มยืนยันหน้า Screen",
                           PV := 5,
                           CV => "Barcode324");
   "M324" := "IEC_Counter_0_DB_351".QU;
   "IEC_Counter_0_DB_1397".CTU(CU := "ยา 325" = 1,
                           R := "Stepper Motor ทำงาน สั่งconveyor เคลื่อที่ไปข้างหน้า" OR "ปุ่มClear",
                           PV := 1);
   "IEC_Counter_0_DB_352".CTUD(CU := ("Expected/Value_All".V = "Expected/Value_All".Expected_325) AND NOT "M325",
                           CD := "IEC_Counter_0_DB_1397".Q AND ("Barcode325" > 0) AND "ปุ่มยืนยันหน้า Screen",
                           PV := 5,
                           CV => "Barcode325");
   "M325" := "IEC_Counter_0_DB_352".QU;
   "IEC_Counter_0_DB_1398".CTU(CU := "ยา 326" = 1,
                           R := "Stepper Motor ทำงาน สั่งconveyor เคลื่อที่ไปข้างหน้า" OR "ปุ่มClear",
                           PV := 1);
   "IEC_Counter_0_DB_353".CTUD(CU := ("Expected/Value_All".V = "Expected/Value_All".Expected_326) AND NOT "M326",
                           CD := "IEC_Counter_0_DB_1398".Q AND ("Barcode326" > 0) AND "ปุ่มยืนยันหน้า Screen",
                           PV := 5,
                           CV => "Barcode326");
   "M326" := "IEC_Counter_0_DB_353".QU;
   "IEC_Counter_0_DB_1399".CTU(CU := "ยา 327" = 1,
                           R := "Stepper Motor ทำงาน สั่งconveyor เคลื่อที่ไปข้างหน้า" OR "ปุ่มClear",
                           PV := 1);
   "IEC_Counter_0_DB_354".CTUD(CU := ("Expected/Value_All".V = "Expected/Value_All".Expected_327) AND NOT "M327",
                           CD := "IEC_Counter_0_DB_1399".Q AND ("Barcode327" > 0) AND "ปุ่มยืนยันหน้า Screen",
                           PV := 5,
                           CV => "Barcode327");
   "M327" := "IEC_Counter_0_DB_354".QU;
   "IEC_Counter_0_DB_1400".CTU(CU := "ยา 328" = 1,
                           R := "Stepper Motor ทำงาน สั่งconveyor เคลื่อที่ไปข้างหน้า" OR "ปุ่มClear",
                           PV := 1);
   "IEC_Counter_0_DB_355".CTUD(CU := ("Expected/Value_All".V = "Expected/Value_All".Expected_328) AND NOT "M328",
                           CD := "IEC_Counter_0_DB_1400".Q AND ("Barcode328" > 0) AND "ปุ่มยืนยันหน้า Screen",
                           PV := 5,
                           CV => "Barcode328");
   "M328" := "IEC_Counter_0_DB_355".QU;
   "IEC_Counter_0_DB_1401".CTU(CU := "ยา 329" = 1,
                           R := "Stepper Motor ทำงาน สั่งconveyor เคลื่อที่ไปข้างหน้า" OR "ปุ่มClear",
                           PV := 1);
   "IEC_Counter_0_DB_356".CTUD(CU := ("Expected/Value_All".V = "Expected/Value_All".Expected_329) AND NOT "M329",
                           CD := "IEC_Counter_0_DB_1401".Q AND ("Barcode329" > 0) AND "ปุ่มยืนยันหน้า Screen",
                           PV := 5,
                           CV => "Barcode329");
   "M329" := "IEC_Counter_0_DB_356".QU;
   "IEC_Counter_0_DB_1402".CTU(CU := "ยา 330" = 1,
                           R := "Stepper Motor ทำงาน สั่งconveyor เคลื่อที่ไปข้างหน้า" OR "ปุ่มClear",
                           PV := 1);
   "IEC_Counter_0_DB_357".CTUD(CU := ("Expected/Value_All".V = "Expected/Value_All".Expected_330) AND NOT "M330",
                           CD := "IEC_Counter_0_DB_1402".Q AND ("Barcode330" > 0) AND "ปุ่มยืนยันหน้า Screen",
                           PV := 5,
                           CV => "Barcode330");
   "M330" := "IEC_Counter_0_DB_357".QU;
   "IEC_Counter_0_DB_1403".CTU(CU := "ยา 331" = 1,
                           R := "Stepper Motor ทำงาน สั่งconveyor เคลื่อที่ไปข้างหน้า" OR "ปุ่มClear",
                           PV := 1);
   "IEC_Counter_0_DB_358".CTUD(CU := ("Expected/Value_All".V = "Expected/Value_All".Expected_331) AND NOT "M331",
                           CD := "IEC_Counter_0_DB_1403".Q AND ("Barcode331" > 0) AND "ปุ่มยืนยันหน้า Screen",
                           PV := 5,
                           CV => "Barcode331");
   "M331" := "IEC_Counter_0_DB_358".QU;
   "IEC_Counter_0_DB_1404".CTU(CU := "ยา 332" = 1,
                           R := "Stepper Motor ทำงาน สั่งconveyor เคลื่อที่ไปข้างหน้า" OR "ปุ่มClear",
                           PV := 1);
   "IEC_Counter_0_DB_359".CTUD(CU := ("Expected/Value_All".V = "Expected/Value_All".Expected_332) AND NOT "M332",
                           CD := "IEC_Counter_0_DB_1404".Q AND ("Barcode332" > 0) AND "ปุ่มยืนยันหน้า Screen",
                           PV := 5,
                           CV => "Barcode332");
   "M332" := "IEC_Counter_0_DB_359".QU;
   "IEC_Counter_0_DB_1405".CTU(CU := "ยา 333" = 1,
                           R := "Stepper Motor ทำงาน สั่งconveyor เคลื่อที่ไปข้างหน้า" OR "ปุ่มClear",
                           PV := 1);
   "IEC_Counter_0_DB_360".CTUD(CU := ("Expected/Value_All".V = "Expected/Value_All".Expected_333) AND NOT "M333",
                           CD := "IEC_Counter_0_DB_1405".Q AND ("Barcode333" > 0) AND "ปุ่มยืนยันหน้า Screen",
                           PV := 5,
                           CV => "Barcode333");
   "M333" := "IEC_Counter_0_DB_360".QU;
   "IEC_Counter_0_DB_1406".CTU(CU := "ยา 334" = 1,
                           R := "Stepper Motor ทำงาน สั่งconveyor เคลื่อที่ไปข้างหน้า" OR "ปุ่มClear",
                           PV := 1);
   "IEC_Counter_0_DB_361".CTUD(CU := ("Expected/Value_All".V = "Expected/Value_All".Expected_334) AND NOT "M334",
                           CD := "IEC_Counter_0_DB_1406".Q AND ("Barcode334" > 0) AND "ปุ่มยืนยันหน้า Screen",
                           PV := 5,
                           CV => "Barcode334");
   "M334" := "IEC_Counter_0_DB_361".QU;
   "IEC_Counter_0_DB_1407".CTU(CU := "ยา 335" = 1,
                           R := "Stepper Motor ทำงาน สั่งconveyor เคลื่อที่ไปข้างหน้า" OR "ปุ่มClear",
                           PV := 1);
   "IEC_Counter_0_DB_362".CTUD(CU := ("Expected/Value_All".V = "Expected/Value_All".Expected_335) AND NOT "M335",
                           CD := "IEC_Counter_0_DB_1407".Q AND ("Barcode335" > 0) AND "ปุ่มยืนยันหน้า Screen",
                           PV := 5,
                           CV => "Barcode335");
   "M335" := "IEC_Counter_0_DB_362".QU;
   "IEC_Counter_0_DB_1408".CTU(CU := "ยา 336" = 1,
                           R := "Stepper Motor ทำงาน สั่งconveyor เคลื่อที่ไปข้างหน้า" OR "ปุ่มClear",
                           PV := 1);
   "IEC_Counter_0_DB_363".CTUD(CU := ("Expected/Value_All".V = "Expected/Value_All".Expected_336) AND NOT "M336",
                           CD := "IEC_Counter_0_DB_1408".Q AND ("Barcode336" > 0) AND "ปุ่มยืนยันหน้า Screen",
                           PV := 5,
                           CV => "Barcode336");
   "M336" := "IEC_Counter_0_DB_363".QU;
   "IEC_Counter_0_DB_1409".CTU(CU := "ยา 337" = 1,
                           R := "Stepper Motor ทำงาน สั่งconveyor เคลื่อที่ไปข้างหน้า" OR "ปุ่มClear",
                           PV := 1);
   "IEC_Counter_0_DB_364".CTUD(CU := ("Expected/Value_All".V = "Expected/Value_All".Expected_337) AND NOT "M337",
                           CD := "IEC_Counter_0_DB_1409".Q AND ("Barcode337" > 0) AND "ปุ่มยืนยันหน้า Screen",
                           PV := 5,
                           CV => "Barcode337");
   "M337" := "IEC_Counter_0_DB_364".QU;
   "IEC_Counter_0_DB_1410".CTU(CU := "ยา 338" = 1,
                           R := "Stepper Motor ทำงาน สั่งconveyor เคลื่อที่ไปข้างหน้า" OR "ปุ่มClear",
                           PV := 1);
   "IEC_Counter_0_DB_365".CTUD(CU := ("Expected/Value_All".V = "Expected/Value_All".Expected_338) AND NOT "M338",
                           CD := "IEC_Counter_0_DB_1410".Q AND ("Barcode338" > 0) AND "ปุ่มยืนยันหน้า Screen",
                           PV := 5,
                           CV => "Barcode338");
   "M338" := "IEC_Counter_0_DB_365".QU;
   "IEC_Counter_0_DB_1411".CTU(CU := "ยา 339" = 1,
                           R := "Stepper Motor ทำงาน สั่งconveyor เคลื่อที่ไปข้างหน้า" OR "ปุ่มClear",
                           PV := 1);
   "IEC_Counter_0_DB_366".CTUD(CU := ("Expected/Value_All".V = "Expected/Value_All".Expected_339) AND NOT "M339",
                           CD := "IEC_Counter_0_DB_1411".Q AND ("Barcode339" > 0) AND "ปุ่มยืนยันหน้า Screen",
                           PV := 5,
                           CV => "Barcode339");
   "M339" := "IEC_Counter_0_DB_366".QU;
   "IEC_Counter_0_DB_1412".CTU(CU := "ยา 340" = 1,
                           R := "Stepper Motor ทำงาน สั่งconveyor เคลื่อที่ไปข้างหน้า" OR "ปุ่มClear",
                           PV := 1);
   "IEC_Counter_0_DB_367".CTUD(CU := ("Expected/Value_All".V = "Expected/Value_All".Expected_340) AND NOT "M340",
                           CD := "IEC_Counter_0_DB_1412".Q AND ("Barcode340" > 0) AND "ปุ่มยืนยันหน้า Screen",
                           PV := 5,
                           CV => "Barcode340");
   "M340" := "IEC_Counter_0_DB_367".QU;
END_REGION

REGION Network 18
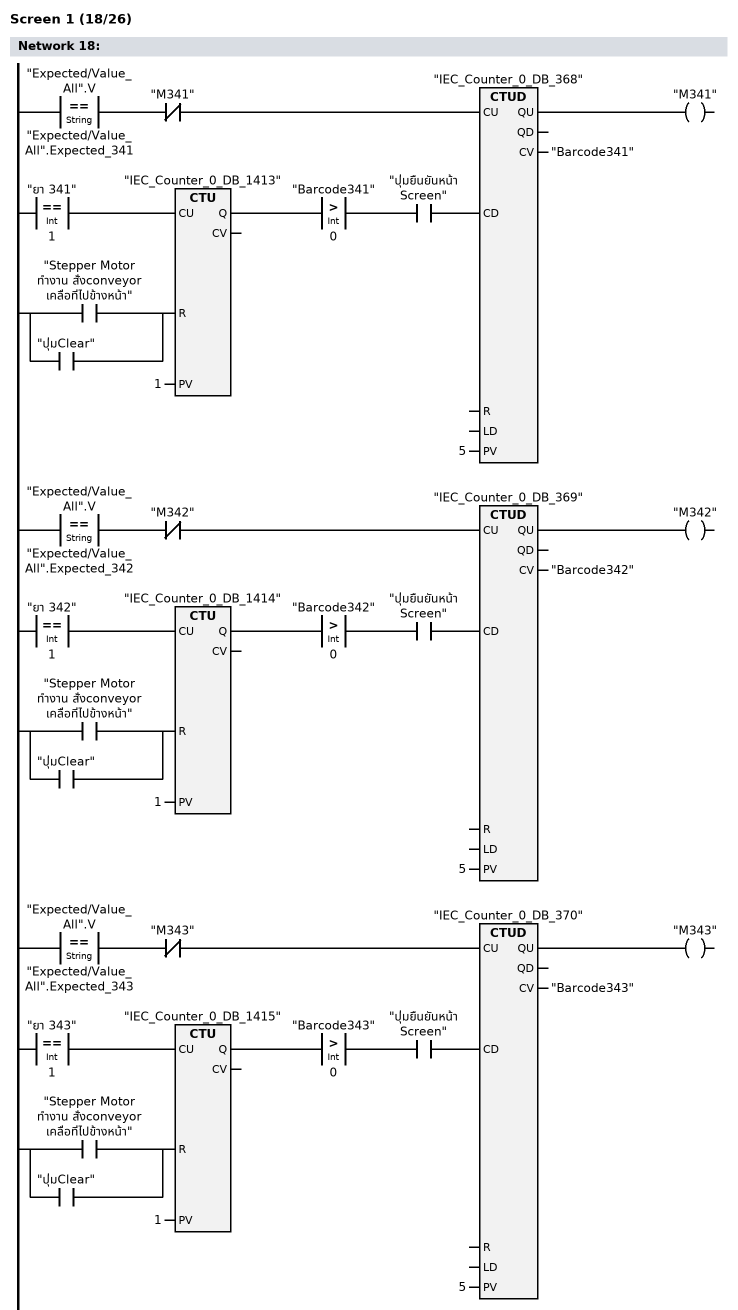
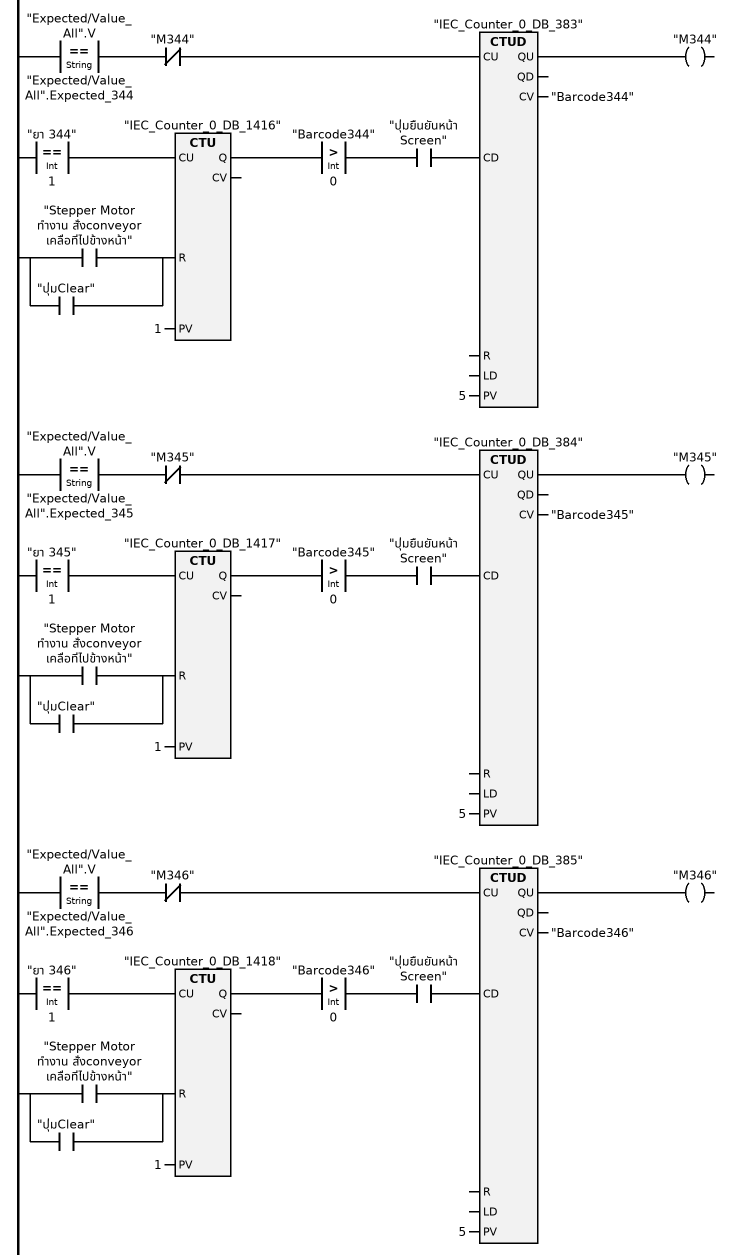
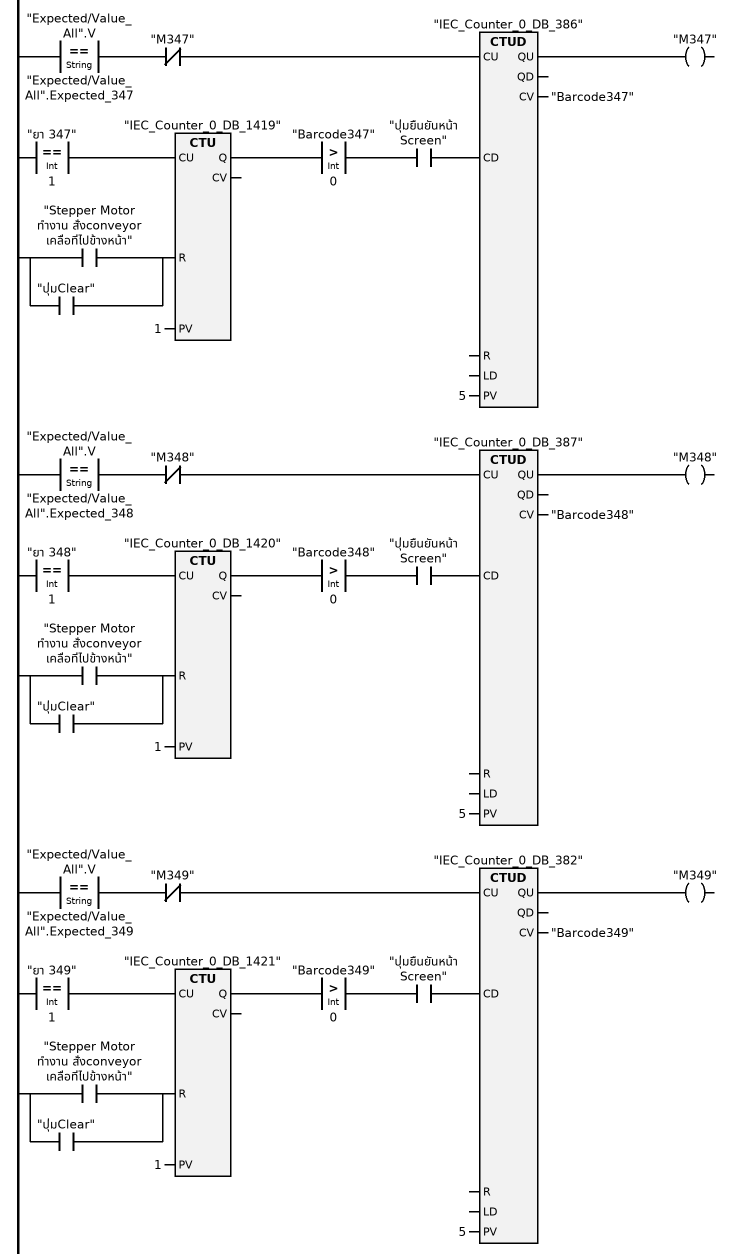
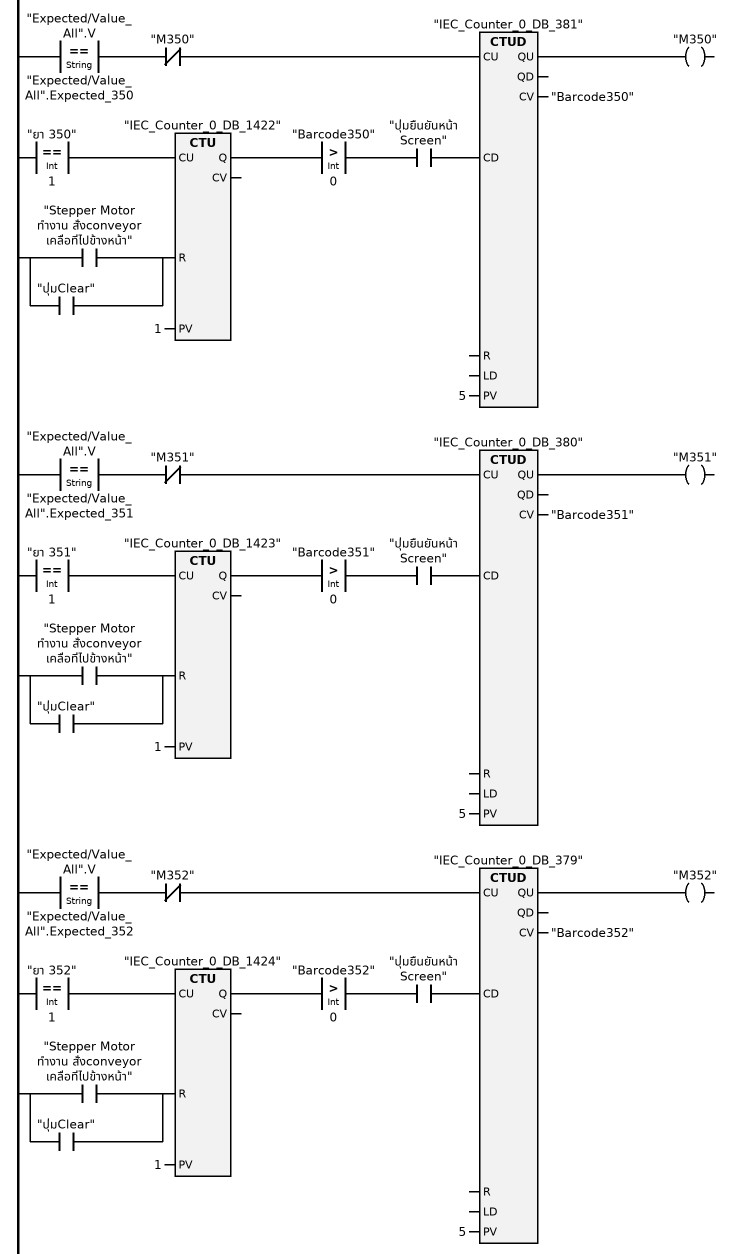
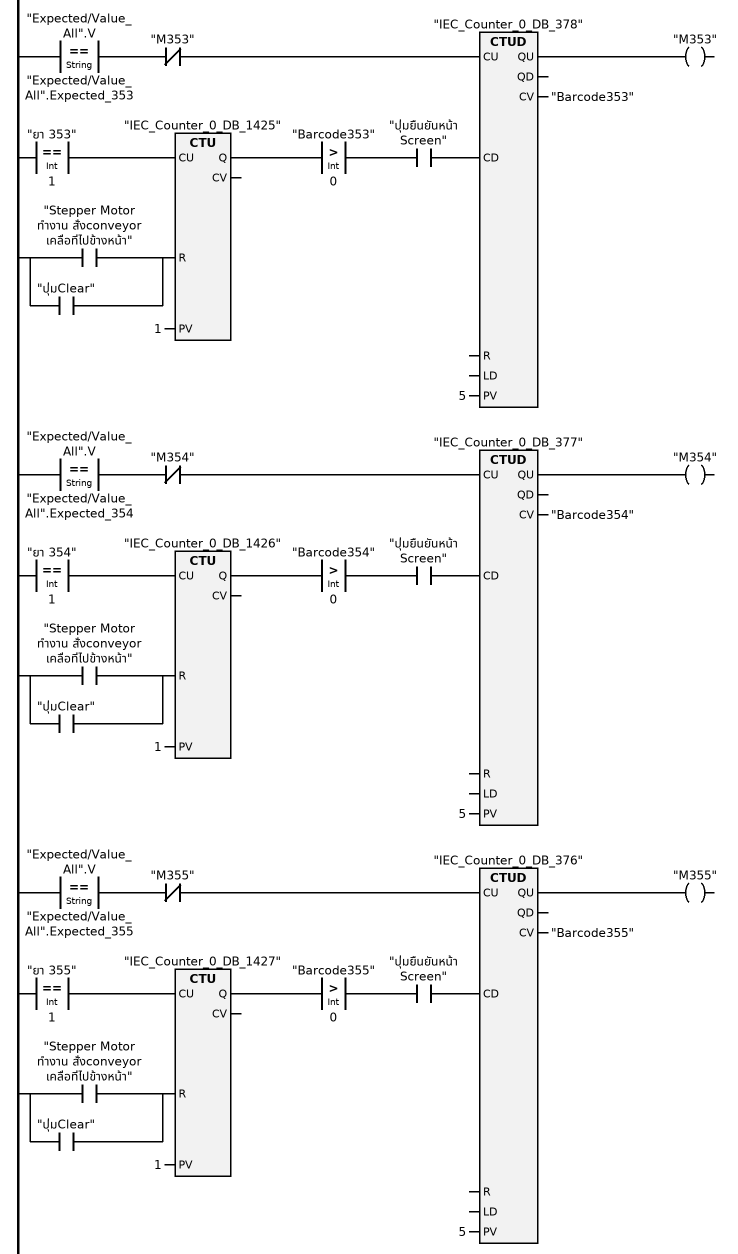
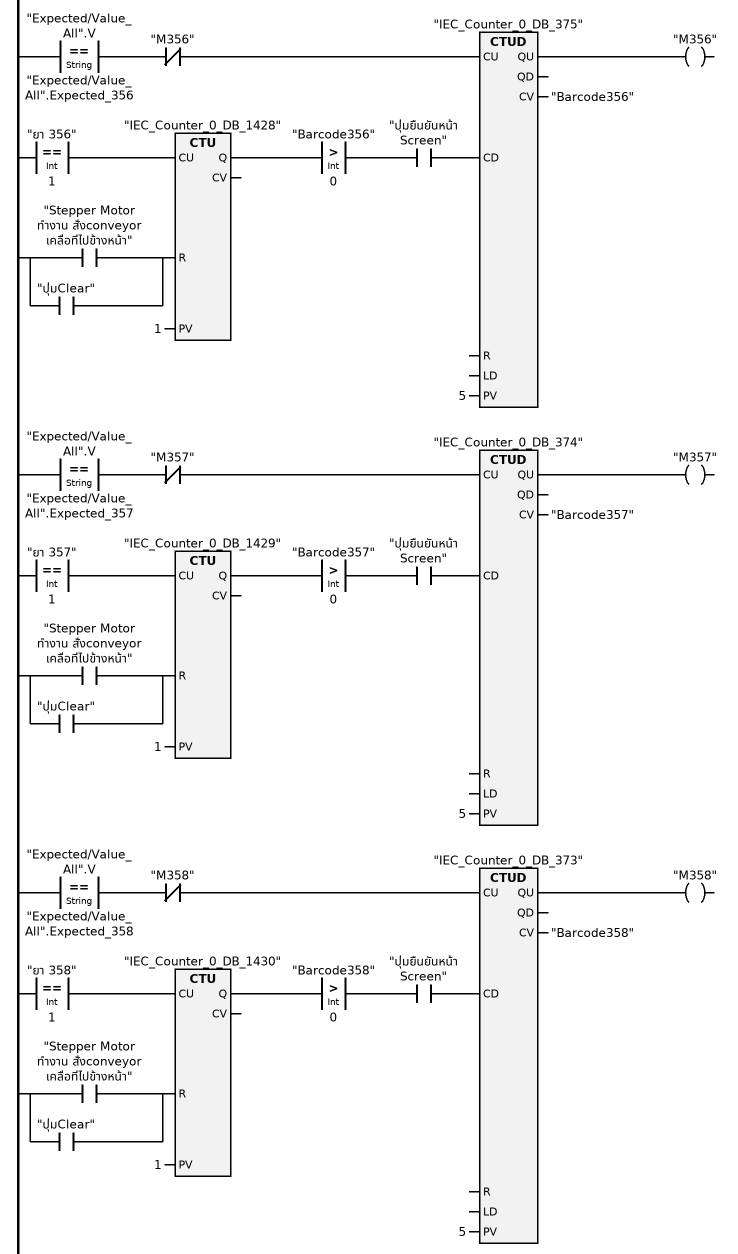
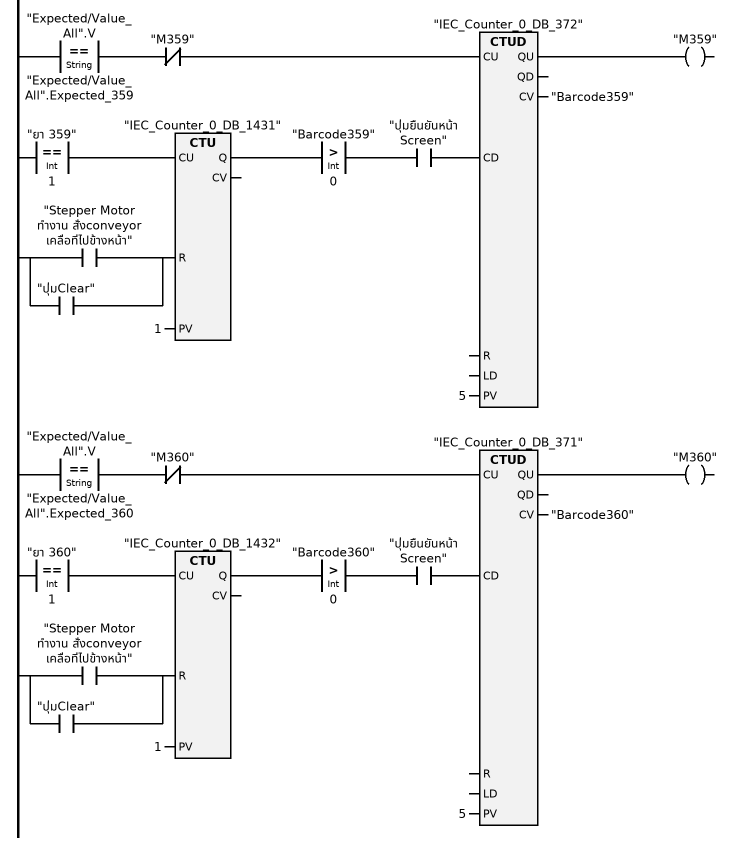
   "IEC_Counter_0_DB_1413".CTU(CU := "ยา 341" = 1,
                           R := "Stepper Motor ทำงาน สั่งconveyor เคลื่อที่ไปข้างหน้า" OR "ปุ่มClear",
                           PV := 1);
   "IEC_Counter_0_DB_368".CTUD(CU := ("Expected/Value_All".V = "Expected/Value_All".Expected_341) AND NOT "M341",
                           CD := "IEC_Counter_0_DB_1413".Q AND ("Barcode341" > 0) AND "ปุ่มยืนยันหน้า Screen",
                           PV := 5,
                           CV => "Barcode341");
   "M341" := "IEC_Counter_0_DB_368".QU;
   "IEC_Counter_0_DB_1414".CTU(CU := "ยา 342" = 1,
                           R := "Stepper Motor ทำงาน สั่งconveyor เคลื่อที่ไปข้างหน้า" OR "ปุ่มClear",
                           PV := 1);
   "IEC_Counter_0_DB_369".CTUD(CU := ("Expected/Value_All".V = "Expected/Value_All".Expected_342) AND NOT "M342",
                           CD := "IEC_Counter_0_DB_1414".Q AND ("Barcode342" > 0) AND "ปุ่มยืนยันหน้า Screen",
                           PV := 5,
                           CV => "Barcode342");
   "M342" := "IEC_Counter_0_DB_369".QU;
   "IEC_Counter_0_DB_1415".CTU(CU := "ยา 343" = 1,
                           R := "Stepper Motor ทำงาน สั่งconveyor เคลื่อที่ไปข้างหน้า" OR "ปุ่มClear",
                           PV := 1);
   "IEC_Counter_0_DB_370".CTUD(CU := ("Expected/Value_All".V = "Expected/Value_All".Expected_343) AND NOT "M343",
                           CD := "IEC_Counter_0_DB_1415".Q AND ("Barcode343" > 0) AND "ปุ่มยืนยันหน้า Screen",
                           PV := 5,
                           CV => "Barcode343");
   "M343" := "IEC_Counter_0_DB_370".QU;
   "IEC_Counter_0_DB_1416".CTU(CU := "ยา 344" = 1,
                           R := "Stepper Motor ทำงาน สั่งconveyor เคลื่อที่ไปข้างหน้า" OR "ปุ่มClear",
                           PV := 1);
   "IEC_Counter_0_DB_383".CTUD(CU := ("Expected/Value_All".V = "Expected/Value_All".Expected_344) AND NOT "M344",
                           CD := "IEC_Counter_0_DB_1416".Q AND ("Barcode344" > 0) AND "ปุ่มยืนยันหน้า Screen",
                           PV := 5,
                           CV => "Barcode344");
   "M344" := "IEC_Counter_0_DB_383".QU;
   "IEC_Counter_0_DB_1417".CTU(CU := "ยา 345" = 1,
                           R := "Stepper Motor ทำงาน สั่งconveyor เคลื่อที่ไปข้างหน้า" OR "ปุ่มClear",
                           PV := 1);
   "IEC_Counter_0_DB_384".CTUD(CU := ("Expected/Value_All".V = "Expected/Value_All".Expected_345) AND NOT "M345",
                           CD := "IEC_Counter_0_DB_1417".Q AND ("Barcode345" > 0) AND "ปุ่มยืนยันหน้า Screen",
                           PV := 5,
                           CV => "Barcode345");
   "M345" := "IEC_Counter_0_DB_384".QU;
   "IEC_Counter_0_DB_1418".CTU(CU := "ยา 346" = 1,
                           R := "Stepper Motor ทำงาน สั่งconveyor เคลื่อที่ไปข้างหน้า" OR "ปุ่มClear",
                           PV := 1);
   "IEC_Counter_0_DB_385".CTUD(CU := ("Expected/Value_All".V = "Expected/Value_All".Expected_346) AND NOT "M346",
                           CD := "IEC_Counter_0_DB_1418".Q AND ("Barcode346" > 0) AND "ปุ่มยืนยันหน้า Screen",
                           PV := 5,
                           CV => "Barcode346");
   "M346" := "IEC_Counter_0_DB_385".QU;
   "IEC_Counter_0_DB_1419".CTU(CU := "ยา 347" = 1,
                           R := "Stepper Motor ทำงาน สั่งconveyor เคลื่อที่ไปข้างหน้า" OR "ปุ่มClear",
                           PV := 1);
   "IEC_Counter_0_DB_386".CTUD(CU := ("Expected/Value_All".V = "Expected/Value_All".Expected_347) AND NOT "M347",
                           CD := "IEC_Counter_0_DB_1419".Q AND ("Barcode347" > 0) AND "ปุ่มยืนยันหน้า Screen",
                           PV := 5,
                           CV => "Barcode347");
   "M347" := "IEC_Counter_0_DB_386".QU;
   "IEC_Counter_0_DB_1420".CTU(CU := "ยา 348" = 1,
                           R := "Stepper Motor ทำงาน สั่งconveyor เคลื่อที่ไปข้างหน้า" OR "ปุ่มClear",
                           PV := 1);
   "IEC_Counter_0_DB_387".CTUD(CU := ("Expected/Value_All".V = "Expected/Value_All".Expected_348) AND NOT "M348",
                           CD := "IEC_Counter_0_DB_1420".Q AND ("Barcode348" > 0) AND "ปุ่มยืนยันหน้า Screen",
                           PV := 5,
                           CV => "Barcode348");
   "M348" := "IEC_Counter_0_DB_387".QU;
   "IEC_Counter_0_DB_1421".CTU(CU := "ยา 349" = 1,
                           R := "Stepper Motor ทำงาน สั่งconveyor เคลื่อที่ไปข้างหน้า" OR "ปุ่มClear",
                           PV := 1);
   "IEC_Counter_0_DB_382".CTUD(CU := ("Expected/Value_All".V = "Expected/Value_All".Expected_349) AND NOT "M349",
                           CD := "IEC_Counter_0_DB_1421".Q AND ("Barcode349" > 0) AND "ปุ่มยืนยันหน้า Screen",
                           PV := 5,
                           CV => "Barcode349");
   "M349" := "IEC_Counter_0_DB_382".QU;
   "IEC_Counter_0_DB_1422".CTU(CU := "ยา 350" = 1,
                           R := "Stepper Motor ทำงาน สั่งconveyor เคลื่อที่ไปข้างหน้า" OR "ปุ่มClear",
                           PV := 1);
   "IEC_Counter_0_DB_381".CTUD(CU := ("Expected/Value_All".V = "Expected/Value_All".Expected_350) AND NOT "M350",
                           CD := "IEC_Counter_0_DB_1422".Q AND ("Barcode350" > 0) AND "ปุ่มยืนยันหน้า Screen",
                           PV := 5,
                           CV => "Barcode350");
   "M350" := "IEC_Counter_0_DB_381".QU;
   "IEC_Counter_0_DB_1423".CTU(CU := "ยา 351" = 1,
                           R := "Stepper Motor ทำงาน สั่งconveyor เคลื่อที่ไปข้างหน้า" OR "ปุ่มClear",
                           PV := 1);
   "IEC_Counter_0_DB_380".CTUD(CU := ("Expected/Value_All".V = "Expected/Value_All".Expected_351) AND NOT "M351",
                           CD := "IEC_Counter_0_DB_1423".Q AND ("Barcode351" > 0) AND "ปุ่มยืนยันหน้า Screen",
                           PV := 5,
                           CV => "Barcode351");
   "M351" := "IEC_Counter_0_DB_380".QU;
   "IEC_Counter_0_DB_1424".CTU(CU := "ยา 352" = 1,
                           R := "Stepper Motor ทำงาน สั่งconveyor เคลื่อที่ไปข้างหน้า" OR "ปุ่มClear",
                           PV := 1);
   "IEC_Counter_0_DB_379".CTUD(CU := ("Expected/Value_All".V = "Expected/Value_All".Expected_352) AND NOT "M352",
                           CD := "IEC_Counter_0_DB_1424".Q AND ("Barcode352" > 0) AND "ปุ่มยืนยันหน้า Screen",
                           PV := 5,
                           CV => "Barcode352");
   "M352" := "IEC_Counter_0_DB_379".QU;
   "IEC_Counter_0_DB_1425".CTU(CU := "ยา 353" = 1,
                           R := "Stepper Motor ทำงาน สั่งconveyor เคลื่อที่ไปข้างหน้า" OR "ปุ่มClear",
                           PV := 1);
   "IEC_Counter_0_DB_378".CTUD(CU := ("Expected/Value_All".V = "Expected/Value_All".Expected_353) AND NOT "M353",
                           CD := "IEC_Counter_0_DB_1425".Q AND ("Barcode353" > 0) AND "ปุ่มยืนยันหน้า Screen",
                           PV := 5,
                           CV => "Barcode353");
   "M353" := "IEC_Counter_0_DB_378".QU;
   "IEC_Counter_0_DB_1426".CTU(CU := "ยา 354" = 1,
                           R := "Stepper Motor ทำงาน สั่งconveyor เคลื่อที่ไปข้างหน้า" OR "ปุ่มClear",
                           PV := 1);
   "IEC_Counter_0_DB_377".CTUD(CU := ("Expected/Value_All".V = "Expected/Value_All".Expected_354) AND NOT "M354",
                           CD := "IEC_Counter_0_DB_1426".Q AND ("Barcode354" > 0) AND "ปุ่มยืนยันหน้า Screen",
                           PV := 5,
                           CV => "Barcode354");
   "M354" := "IEC_Counter_0_DB_377".QU;
   "IEC_Counter_0_DB_1427".CTU(CU := "ยา 355" = 1,
                           R := "Stepper Motor ทำงาน สั่งconveyor เคลื่อที่ไปข้างหน้า" OR "ปุ่มClear",
                           PV := 1);
   "IEC_Counter_0_DB_376".CTUD(CU := ("Expected/Value_All".V = "Expected/Value_All".Expected_355) AND NOT "M355",
                           CD := "IEC_Counter_0_DB_1427".Q AND ("Barcode355" > 0) AND "ปุ่มยืนยันหน้า Screen",
                           PV := 5,
                           CV => "Barcode355");
   "M355" := "IEC_Counter_0_DB_376".QU;
   "IEC_Counter_0_DB_1428".CTU(CU := "ยา 356" = 1,
                           R := "Stepper Motor ทำงาน สั่งconveyor เคลื่อที่ไปข้างหน้า" OR "ปุ่มClear",
                           PV := 1);
   "IEC_Counter_0_DB_375".CTUD(CU := ("Expected/Value_All".V = "Expected/Value_All".Expected_356) AND NOT "M356",
                           CD := "IEC_Counter_0_DB_1428".Q AND ("Barcode356" > 0) AND "ปุ่มยืนยันหน้า Screen",
                           PV := 5,
                           CV => "Barcode356");
   "M356" := "IEC_Counter_0_DB_375".QU;
   "IEC_Counter_0_DB_1429".CTU(CU := "ยา 357" = 1,
                           R := "Stepper Motor ทำงาน สั่งconveyor เคลื่อที่ไปข้างหน้า" OR "ปุ่มClear",
                           PV := 1);
   "IEC_Counter_0_DB_374".CTUD(CU := ("Expected/Value_All".V = "Expected/Value_All".Expected_357) AND NOT "M357",
                           CD := "IEC_Counter_0_DB_1429".Q AND ("Barcode357" > 0) AND "ปุ่มยืนยันหน้า Screen",
                           PV := 5,
                           CV => "Barcode357");
   "M357" := "IEC_Counter_0_DB_374".QU;
   "IEC_Counter_0_DB_1430".CTU(CU := "ยา 358" = 1,
                           R := "Stepper Motor ทำงาน สั่งconveyor เคลื่อที่ไปข้างหน้า" OR "ปุ่มClear",
                           PV := 1);
   "IEC_Counter_0_DB_373".CTUD(CU := ("Expected/Value_All".V = "Expected/Value_All".Expected_358) AND NOT "M358",
                           CD := "IEC_Counter_0_DB_1430".Q AND ("Barcode358" > 0) AND "ปุ่มยืนยันหน้า Screen",
                           PV := 5,
                           CV => "Barcode358");
   "M358" := "IEC_Counter_0_DB_373".QU;
   "IEC_Counter_0_DB_1431".CTU(CU := "ยา 359" = 1,
                           R := "Stepper Motor ทำงาน สั่งconveyor เคลื่อที่ไปข้างหน้า" OR "ปุ่มClear",
                           PV := 1);
   "IEC_Counter_0_DB_372".CTUD(CU := ("Expected/Value_All".V = "Expected/Value_All".Expected_359) AND NOT "M359",
                           CD := "IEC_Counter_0_DB_1431".Q AND ("Barcode359" > 0) AND "ปุ่มยืนยันหน้า Screen",
                           PV := 5,
                           CV => "Barcode359");
   "M359" := "IEC_Counter_0_DB_372".QU;
   "IEC_Counter_0_DB_1432".CTU(CU := "ยา 360" = 1,
                           R := "Stepper Motor ทำงาน สั่งconveyor เคลื่อที่ไปข้างหน้า" OR "ปุ่มClear",
                           PV := 1);
   "IEC_Counter_0_DB_371".CTUD(CU := ("Expected/Value_All".V = "Expected/Value_All".Expected_360) AND NOT "M360",
                           CD := "IEC_Counter_0_DB_1432".Q AND ("Barcode360" > 0) AND "ปุ่มยืนยันหน้า Screen",
                           PV := 5,
                           CV => "Barcode360");
   "M360" := "IEC_Counter_0_DB_371".QU;
END_REGION

REGION Network 19
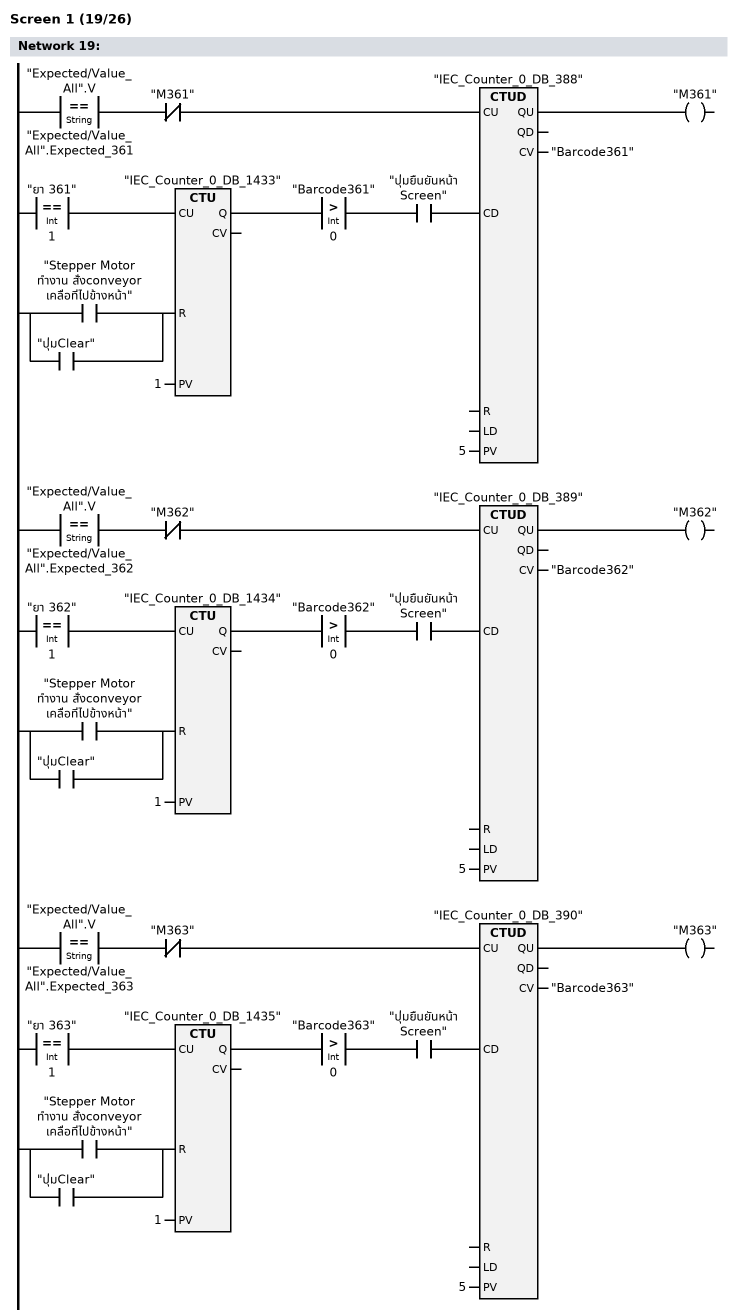
